(* IEC 61131-3 sources: daoli-st-library/DL_Process (part 14) *)

(* ---- FC_DL_LyoCollapseTempMarginCalc.st ---- *)
(*
  Name: FC_DL_LyoCollapseTempMarginCalc
  Category: DL_Process
  Version: 1.0.0
  Round: R91 / 2026-11-25
  开源溯源：clean-room 自研（族 制药冻干真空冷冻干燥，ST 开源生态实测 0 命中，无外部代码引入）
  功能：1) 塌陷温度裕度 = 塌陷温度 − 制品温度，即 fMarginK = fCollapseC − fProductC，
           裕度为正表示制品温度仍低于塌陷温度（安全侧），为负表示已越过塌陷边界。
        2) 裕度分级（nGrade）：0 = 合格（裕度 >= fMarginWarnK），1 = 预警（fMarginMinK <= 裕度 < fMarginWarnK），
           2 = 不足（裕度 < fMarginMinK），分级判据全部对原始裕度做，钳制只作用于输出数值。
        3) 冰点约束：制品温度必须低于冰点 fIcePointC，否则一次干燥已进入液态（融冰），
           输出 xAboveIce 供上层立即降温或转二次干燥。
  边界条件：1) 非有限值闸：五路实值入参先过 NOT(x > -DL_BIG AND x < DL_BIG)，同时拦 NaN 与 Inf，
           命中即闸断实值通路（裕度强制 0.0 且置分级 2 = 不足），不得只置标志（R19）。
        2) 阈值域闸：分级阈值须满足 fMarginMinK < fMarginWarnK（否则两级判据区间为空、分级恒失效），
           越域判无效并把 nGrade 置 2（保守侧）。
        3) 温度域闸：三路温度必须落在 [-DL_T_SPAN, +DL_T_SPAN] 内，越域判无效（量级异常）。
        4) 判据取原始值（R24）：分级与冰点判定使用原始入参，不先把温度夹到工艺带再判。
        5) 物理域钳制：裕度钳到 [-DL_MARGIN_SPAN, +DL_MARGIN_SPAN]，避免极端值污染显示与趋势。
        6) 纯函数无状态：分级不做迟滞，防抖与联锁延时由搁板温控 FB 承担。
  量纲自证：fMarginK = (degC) − (degC) = (K)；与 fMarginMinK / fMarginWarnK 同为温差点量纲 [K]，
           可与温差阈值直接比较；nGrade 为无量纲等级 [level]。
  修订历史 Revision :
    2026-11-25  v1.0.0  R91 首版
*)

FUNCTION FC_DL_LyoCollapseTempMarginCalc : BOOL
VAR_INPUT
    fProductC        : REAL;   // 制品（瓶内）温度 [degC] / Product temperature inside the vial [degC]
    fCollapseC       : REAL;   // 配方给出的塌陷温度 [degC] / Formulation collapse temperature [degC]
    fIcePointC       : REAL;   // 配方给出的冰点 [degC] / Formulation ice point [degC]
    fMarginMinK      : REAL;   // 裕度不足阈值（低于即判不足）[K] / Margin insufficient threshold [K]
    fMarginWarnK     : REAL;   // 裕度预警阈值（低于即判预警）[K] / Margin warning threshold [K]
END_VAR
VAR_OUTPUT
    fMarginK         : REAL;   // 塌陷温度裕度 [K] / Collapse temperature margin [K]
    nGrade           : INT;    // 裕度分级 0=合格 1=预警 2=不足 [level] / Margin grade 0/1/2 [level]
    xMarginLow       : BOOL;   // 裕度不足标志（< 下限）[bool] / Margin insufficient flag [bool]
    xAboveIce        : BOOL;   // 制品温度高于冰点标志 [bool] / Product above ice point flag [bool]
    xValid           : BOOL;   // 计算有效标志 [bool] / Calculation valid flag [bool]
END_VAR
VAR
    _fMarginRawK     : REAL;   // 钳制前的原始裕度 [K] / Raw margin before limiting [K]
END_VAR
VAR CONSTANT
    DL_BIG           : REAL := 1.0E12;    // 非有限值闸量级上限 [-] / Finiteness gate magnitude [-]
    DL_EPS           : REAL := 1.0E-9;    // 数值零闸阈值 [-] / Numeric zero gate threshold [-]
    DL_T_SPAN        : REAL := 300.0;     // 温度量级闸跨度 [degC] / Temperature magnitude gate span [degC]
    DL_MARGIN_SPAN   : REAL := 200.0;     // 裕度钳制跨度 [K] / Margin clamp span [K]
    DL_GRADE_OK      : INT := 0;          // 分级：合格 [level] / Grade: acceptable [level]
    DL_GRADE_WARN    : INT := 1;          // 分级：预警 [level] / Grade: warning [level]
    DL_GRADE_BAD     : INT := 2;          // 分级：不足 [level] / Grade: insufficient [level]
END_VAR

(* —— 段 1：非有限值闸（R19：闸断实值通路；失效侧分级置不足） —— *)
IF NOT (fProductC > -DL_BIG AND fProductC < DL_BIG)
   OR NOT (fCollapseC > -DL_BIG AND fCollapseC < DL_BIG)
   OR NOT (fIcePointC > -DL_BIG AND fIcePointC < DL_BIG)
   OR NOT (fMarginMinK > -DL_BIG AND fMarginMinK < DL_BIG)
   OR NOT (fMarginWarnK > -DL_BIG AND fMarginWarnK < DL_BIG) THEN
    fMarginK := 0.0;                        // 输出强制 0.0，切断污染源 / Force zero, cut polluted path
    nGrade := DL_GRADE_BAD;                 // 失效侧按不足处理（保守侧）/ Treat as insufficient when invalid
    xMarginLow := TRUE;                     // 失效侧不足位置真（保守侧）/ Insufficient flag true when invalid
    xAboveIce := FALSE;                     // 失效侧冰点位保持假 / Ice-point flag stays false
    xValid := FALSE;                        // 有效位清零 / Validity cleared
    FC_DL_LyoCollapseTempMarginCalc := FALSE;   // 返回码与有效位同源 / Return mirrors validity
    RETURN;                                 // 立即退出 / Immediate exit
END_IF

(* —— 段 2：主算式（不钳制，先出原始值供段 3 判据使用，R24） —— *)
_fMarginRawK := fCollapseC - fProductC;                                           // 塌陷温度裕度 [K]

(* —— 段 3：判据与分级（全部取原始值；单点 BOOL 聚合避免多处赋 FALSE 覆盖） —— *)
xMarginLow := (_fMarginRawK < fMarginMinK);                                       // 裕度不足
xAboveIce := (fProductC > fIcePointC);                                            // 已融冰（高于冰点）
xValid := (fMarginMinK < fMarginWarnK)                                            // 分级阈值必须有效（min < warn）
          AND (ABS(fProductC) <= DL_T_SPAN)                                       // 温度量级闸
          AND (ABS(fCollapseC) <= DL_T_SPAN)
          AND (ABS(fIcePointC) <= DL_T_SPAN)
          AND (fCollapseC > fIcePointC);                                          // 塌陷温度须高于冰点（物理约束）

IF NOT xValid THEN
    nGrade := DL_GRADE_BAD;                 // 参数非法：按不足处理（保守侧）
ELSIF _fMarginRawK >= fMarginWarnK THEN
    nGrade := DL_GRADE_OK;                  // 裕度充足
ELSIF _fMarginRawK >= fMarginMinK THEN
    nGrade := DL_GRADE_WARN;                // 预警带
ELSE
    nGrade := DL_GRADE_BAD;                 // 不足
END_IF

(* —— 段 4：输出单点写盘（钳制到物理域内，分级已在段 3 定案） —— *)
fMarginK := LIMIT(-DL_MARGIN_SPAN, _fMarginRawK, DL_MARGIN_SPAN);                  // 裕度钳到物理域 [K]
FC_DL_LyoCollapseTempMarginCalc := xValid;                                        // 返回码：TRUE = 计算可信

END_FUNCTION

(* ---- FC_DL_LyoIceVaporPressureCalc.st ---- *)
(*
  Name: FC_DL_LyoIceVaporPressureCalc
  Category: DL_Process
  Version: 1.0.0
  Round: R91 / 2026-11-25
  开源溯源：clean-room 自研（族 制药冻干真空冷冻干燥，ST 开源生态实测 0 命中，无外部代码引入）
  功能：1) 冰面饱和蒸气压按 Magnus 型 Goff-Gratch 简化式求解：
           p_ice = 611.15 * EXP(22.452 * T / (272.55 + T))，T 为冰面温度 [degC]，
           611.15 为 0 degC 时冰面饱和蒸气压 [Pa]，22.452 与 272.55 为冰相经验常数。
           该式在 -60 ~ 0 degC 内相对误差小于 1 %，是冻干一次干燥压力设定的标准依据。
        2) 派生输出过冷度裕量 fSubcoolK = 0.0 − T，即离冰点的距离；
           冻干工艺要求制品温度始终低于冰点，裕量为负意味着已融冰（塌陷前兆）。
        3) 温度域校验：温度必须落在 [DL_T_LO, DL_T_HI] = [-60.0, 0.0] degC 内，
           越域只置 xDomainOk = FALSE 而数值钳到域内输出，因为经验常数在域外已失效。
  边界条件：1) 非有限值闸：温度入参先过 NOT(x > -DL_BIG AND x < DL_BIG)，同时拦 NaN 与 Inf，
           命中即闸断实值通路（fPressurePa 与 fSubcoolK 强制 0.0），不得只置标志（R19）。
        2) 分母零闸：经验式分母 272.55 + T 在 T = -272.55 degC 处为零，
           本件温度域下限 -60 degC 远高于该点，但仍显式校验 |272.55 + T| > DL_EPS，
           防止越域调用（下游误传开尔文值）导致除零。
        3) 指数溢出闸：指数 22.452*T/(272.55+T) 在接近 -272.55 时发散，
           计算前用温度域闸先拦截，绝不让 EXP 收到发散指数（EXP 溢出为 Inf 会穿透下游）。
        4) 判据取原始值（R24）：温度越域判定使用原始入参 fTempC，不对其先钳制再判。
        5) 物理域钳制：气压钳 0.0 ~ DL_P_HI_PA；过冷度钳到 [-DL_T_HI_SPAN, +DL_T_HI_SPAN]。
        6) 纯函数无状态：不做滤波，测点噪声抑制由下游一阶滤波件承担。
  量纲自证：T [degC] 代入经验式时以温差形式参与（degC 与 K 的差值尺度相同），
           22.452*T/(272.55+T) = (无因次)，故 EXP 的自变量无因次；
           p_ice = (Pa) * (无因次) = Pa，量纲合法。
  修订历史 Revision :
    2026-11-25  v1.0.0  R91 首版
*)

FUNCTION FC_DL_LyoIceVaporPressureCalc : BOOL
VAR_INPUT
    fTempC           : REAL;   // 冰面温度 [degC] / Ice surface temperature [degC]
END_VAR
VAR_OUTPUT
    fPressurePa      : REAL;   // 冰面饱和蒸气压 [Pa] / Ice surface saturation vapour pressure [Pa]
    fSubcoolK        : REAL;   // 距冰点的过冷度裕量 [K] / Subcooling margin below the ice point [K]
    xDomainOk        : BOOL;   // 温度在经验式有效域内 [bool] / Temperature within the valid domain [bool]
    xValid           : BOOL;   // 计算有效标志 [bool] / Calculation valid flag [bool]
END_VAR
VAR
    _fDenomK         : REAL;   // 经验式分母（272.55 + T）[K] / Empirical denominator, 272.55 + T [K]
    _fExpo           : REAL;   // 经验式指数（无因次）[-] / Empirical exponent, dimensionless [-]
    _fPressRawPa     : REAL;   // 钳制前的原始气压 [Pa] / Raw pressure before limiting [Pa]
    _fTempUseC       : REAL;   // 域钳制后参与计算的温度 [degC] / Temperature used after domain clamping [degC]
END_VAR
VAR CONSTANT
    DL_EPS           : REAL := 1.0E-9;    // 数值零闸阈值 [-] / Numeric zero gate threshold [-]
    DL_BIG           : REAL := 1.0E12;    // 非有限值闸量级上限 [-] / Finiteness gate magnitude [-]
    DL_T_LO          : REAL := -60.0;     // 经验式有效温度下限 [degC] / Valid temperature low bound [degC]
    DL_T_HI          : REAL := 0.0;       // 经验式有效温度上限（冰点）[degC] / Valid temperature high, ice point [degC]
    DL_P0_PA         : REAL := 611.15;    // 0 degC 冰面饱和蒸气压 [Pa] / Ice saturation pressure at 0 degC [Pa]
    DL_COEF_A        : REAL := 22.452;    // 冰相经验常数 A（无因次）[-] / Ice-phase empirical constant A [-]
    DL_COEF_B        : REAL := 272.55;    // 冰相经验常数 B [K] / Ice-phase empirical constant B [K]
    DL_P_HI_PA       : REAL := 700.0;     // 气压物理上限（略高于 0 degC 冰面值）[Pa] / Pressure upper bound [Pa]
    DL_MARGIN_SPAN   : REAL := 200.0;     // 过冷度裕量钳制跨度 [K] / Subcooling margin clamp span [K]
END_VAR

(* —— 段 1：非有限值闸（R19：闸断实值通路） —— *)
IF NOT (fTempC > -DL_BIG AND fTempC < DL_BIG) THEN
    fPressurePa := 0.0;                     // 输出强制 0.0，切断污染源 / Force zero, cut polluted path
    fSubcoolK := 0.0;                       // 裕量强制 0.0 / Margin forced to zero
    xDomainOk := FALSE;                     // 域位清零 / Domain flag cleared
    xValid := FALSE;                        // 有效位清零 / Validity cleared
    FC_DL_LyoIceVaporPressureCalc := FALSE; // 返回码与有效位同源 / Return mirrors validity
    RETURN;                                 // 立即退出 / Immediate exit
END_IF

(* —— 段 2：判据取原始值（R24：先判域，再钳制，禁先钳后判） —— *)
xDomainOk := (fTempC >= DL_T_LO) AND (fTempC <= DL_T_HI);

(* —— 段 3：域钳制后参与计算（经验常数在域外失效，绝不让 EXP 收到发散指数） —— *)
_fTempUseC := LIMIT(DL_T_LO, fTempC, DL_T_HI);                          // 温度钳到有效域 [degC]
_fDenomK := DL_COEF_B + _fTempUseC;                                     // 经验式分母 [K]

(* —— 段 4：分母零闸（防越域调用传开尔文值导致除零，R4） —— *)
IF ABS(_fDenomK) <= DL_EPS THEN
    fPressurePa := 0.0;                     // 分母为零即不可算 / No denominator, no result
    fSubcoolK := 0.0;                       // 裕量不可算 / Margin not computable
    xDomainOk := FALSE;                     // 判域外 / Out of domain
    xValid := FALSE;                        // 判无效 / Invalid
    FC_DL_LyoIceVaporPressureCalc := FALSE; // 返回码同步 / Return synchronised
    RETURN;                                 // 提前退出 / Early exit
END_IF

(* —— 段 5：主算式（Goff-Gratch 简化式，指数自变量已由段 3 钳制保证有界） —— *)
_fExpo := DL_COEF_A * _fTempUseC / _fDenomK;                            // 指数（无因次）[-]
_fPressRawPa := DL_P0_PA * EXP(_fExpo);                                 // 冰面饱和蒸气压 [Pa]
fSubcoolK := LIMIT(-DL_MARGIN_SPAN, DL_T_HI - _fTempUseC, DL_MARGIN_SPAN);   // 过冷度裕量 [K]

(* —— 段 6：输出单点写盘（气压钳制到物理域；有限性已由段 1 保证） —— *)
fPressurePa := LIMIT(0.0, _fPressRawPa, DL_P_HI_PA);                    // 气压钳 0..物理上限 [Pa]
xValid := xDomainOk AND (fPressurePa > 0.0);                            // 域内且有正压才算有效
FC_DL_LyoIceVaporPressureCalc := xValid;                                // 返回码：TRUE = 计算可信

END_FUNCTION

(* ---- FC_DL_LyoPrimaryDryingTimeCalc.st ---- *)
(*
  Name: FC_DL_LyoPrimaryDryingTimeCalc
  Category: DL_Process
  Version: 1.0.0
  Round: R91 / 2026-11-25
  开源溯源：clean-room 自研（族 制药冻干真空冷冻干燥，ST 开源生态实测 0 命中，无外部代码引入）
  功能：1) 一次干燥时间按「可去除水量 / 升华速率」估算：
           可去除水量 W = 装量质量 * (初始含水率 − 目标含水率) / 100，单位 kg；
           时间 t = W / rate，单位 h；rate 为该批量的实测升华速率 [kg/h]。
        2) 水量守恒校验：目标含水率必须低于初始含水率，否则水量为负（配方错），
           判无效而不取绝对值 —— 负水量意味着「越干越湿」的错误配方。
        3) 收敛判据：估算时间超过 fMaxTimeH（工艺允许最长一次干燥时间）时置 xNotConverge，
           表示按当前速率无法在允许时间内达到目标含水率，需提高搁板温度或降低装量。
  边界条件：1) 非有限值闸：五路实值入参先过 NOT(x > -DL_BIG AND x < DL_BIG)，同时拦 NaN 与 Inf，
           命中即闸断实值通路（时间与水量强制 0.0），不得只置标志（R19）。
        2) 速率零闸：升华速率 fRateKgh 必须 > DL_EPS（时间式的分母），否则判无效并清零，
           不得输出「无穷长时间」这种不可执行值。
        3) 含水率域闸：初始与目标含水率必须落在 [0.0, 100.0] % 内，
           装量质量须 > DL_EPS；任一越域判无效，不做钳制。
        4) 判据取原始值（R24）：不收敛判定使用钳制前的 _fTimeRawH，不得先钳再判。
        5) 物理域钳制：时间钳 0.0 ~ DL_TIME_HI_H；水量钳 0.0 ~ 装量质量（水量不可能大于装量）。
        6) 纯函数无状态：不累计已干燥时间，累计与阶段切换由干燥序 FB 承担。
  量纲自证：W = (kg) * (无因次百分数/100) = kg；
           t = (kg)/(kg/h) = h，与 fMaxTimeH 同量纲 [h]，可直接比较。
  修订历史 Revision :
    2026-11-25  v1.0.0  R91 首版
*)

FUNCTION FC_DL_LyoPrimaryDryingTimeCalc : BOOL
VAR_INPUT
    fFillMassKg      : REAL;   // 单批装量质量 [kg] / Batch fill mass [kg]
    fInitMoistPct    : REAL;   // 初始含水率 [%] / Initial moisture content [%]
    fTargetMoistPct  : REAL;   // 目标含水率 [%] / Target moisture content [%]
    fRateKgh         : REAL;   // 该批量实测升华速率 [kg/h] / Measured batch sublimation rate [kg/h]
    fMaxTimeH        : REAL;   // 工艺允许最长一次干燥时间 [h] / Permitted maximum primary drying time [h]
END_VAR
VAR_OUTPUT
    fTimeH           : REAL;   // 一次干燥估算时间 [h] / Estimated primary drying time [h]
    fWaterKg         : REAL;   // 需去除水量 [kg] / Water mass to be removed [kg]
    xNotConverge     : BOOL;   // 超允许时间标志（不收敛）[bool] / Non-convergence flag [bool]
    xValid           : BOOL;   // 计算有效标志 [bool] / Calculation valid flag [bool]
END_VAR
VAR
    _fWaterRawKg     : REAL;   // 钳制前的原始水量 [kg] / Raw water mass before limiting [kg]
    _fTimeRawH       : REAL;   // 钳制前的原始时间 [h] / Raw time before limiting [h]
END_VAR
VAR CONSTANT
    DL_EPS           : REAL := 1.0E-9;    // 数值零闸阈值 [-] / Numeric zero gate threshold [-]
    DL_BIG           : REAL := 1.0E12;    // 非有限值闸量级上限 [-] / Finiteness gate magnitude [-]
    DL_PCT           : REAL := 100.0;     // 百分比换算因子（含水率分母）[%] / Percent conversion factor [%]
    DL_PCT_HI        : REAL := 100.0;     // 含水率物理上限 [%] / Moisture content upper bound [%]
    DL_TIME_HI_H     : REAL := 10000.0;   // 时间物理上限 [h] / Time physical upper bound [h]
END_VAR

(* —— 段 1：非有限值闸（R19：闸断实值通路） —— *)
IF NOT (fFillMassKg > -DL_BIG AND fFillMassKg < DL_BIG)
   OR NOT (fInitMoistPct > -DL_BIG AND fInitMoistPct < DL_BIG)
   OR NOT (fTargetMoistPct > -DL_BIG AND fTargetMoistPct < DL_BIG)
   OR NOT (fRateKgh > -DL_BIG AND fRateKgh < DL_BIG)
   OR NOT (fMaxTimeH > -DL_BIG AND fMaxTimeH < DL_BIG) THEN
    fTimeH := 0.0;                          // 输出强制 0.0，切断污染源 / Force zero, cut polluted path
    fWaterKg := 0.0;                        // 水量强制 0.0 / Water mass forced to zero
    xNotConverge := TRUE;                   // 失效侧按不收敛处理（安全侧）/ Treat as non-converged when invalid
    xValid := FALSE;                        // 有效位清零 / Validity cleared
    FC_DL_LyoPrimaryDryingTimeCalc := FALSE;   // 返回码与有效位同源 / Return mirrors validity
    RETURN;                                 // 立即退出 / Immediate exit
END_IF

(* —— 段 2：分母零闸与域闸（时间式分母为速率；含水率须在 0~100 %） —— *)
IF (fRateKgh <= DL_EPS)                                           // 速率不可为零
   OR (fFillMassKg <= DL_EPS)                                     // 装量不可为零
   OR (fInitMoistPct < 0.0)                                       // 含水率不得为负
   OR (fInitMoistPct > DL_PCT_HI)                                 // 含水率不得超 100 %
   OR (fTargetMoistPct < 0.0)                                     // 目标含水率不得为负
   OR (fTargetMoistPct > DL_PCT_HI)                               // 目标含水率不得超 100 %
   OR (fMaxTimeH <= DL_EPS) THEN                                  // 允许时间必须已组态
    fTimeH := 0.0;                          // 参数不可用即无时间 / No parameter, no time
    fWaterKg := 0.0;                        // 水量不可算 / Water mass not computable
    xNotConverge := TRUE;                   // 按不收敛处理 / Treat as non-converged
    xValid := FALSE;                        // 判无效 / Invalid
    FC_DL_LyoPrimaryDryingTimeCalc := FALSE;   // 返回码同步 / Return synchronised
    RETURN;                                 // 提前退出 / Early exit
END_IF

(* —— 段 3：主算式（不钳制，先出原始值供段 4 判据使用，R24） —— *)
_fWaterRawKg := fFillMassKg * (fInitMoistPct - fTargetMoistPct) / DL_PCT;          // 需去除水量 [kg]
_fTimeRawH := _fWaterRawKg / fRateKgh;                                            // 估算时间 [h]

(* —— 段 4：判据（取原始值；单点 BOOL 聚合避免多处赋 FALSE 覆盖） —— *)
xNotConverge := (_fTimeRawH > fMaxTimeH);                                         // 超允许时间：不收敛
xValid := (_fWaterRawKg >= 0.0)                                                   // 水量不得为负（配方方向固定）
          AND (_fTimeRawH >= 0.0)                                                 // 时间不得为负
          AND (fMaxTimeH <= DL_TIME_HI_H)                                         // 允许时间不得超物理上限
          AND (fInitMoistPct > fTargetMoistPct);                                  // 初始必须高于目标（方向固定）

(* —— 段 5：输出单点写盘（钳制到物理域内，判定结果已在段 4 定案） —— *)
fWaterKg := LIMIT(0.0, _fWaterRawKg, fFillMassKg);                                // 水量钳 0..装量 [kg]
fTimeH := LIMIT(0.0, _fTimeRawH, DL_TIME_HI_H);                                   // 时间钳 0..物理上限 [h]
FC_DL_LyoPrimaryDryingTimeCalc := xValid;                                         // 返回码：TRUE = 计算可信

END_FUNCTION

(* ---- FC_DL_LyoResidualMoistureCalc.st ---- *)
(*
  Name: FC_DL_LyoResidualMoistureCalc
  Category: DL_Process
  Version: 1.0.0
  Round: R91 / 2026-11-25
  开源溯源：clean-room 自研（族 制药冻干真空冷冻干燥，ST 开源生态实测 0 命中，无外部代码引入）
  功能：1) 残余水分估算按「压力升速率法」：一次干燥末期关闭隔离阀，测腔内压力升幅与时间，
           升压速率 r = dP / t [mbar/s]；残余水分与升压速率近似成正比，并用干重比归一：
           W_res% = coef * r / ratio，coef 为经方法学验证的标定系数 [%*s/mbar]，
           ratio 为干物质质量占比 [kg/kg]（干重比），用于把腔体自由水折算到制品含湿量。
        2) 合格判据：残余水分 <= fSpecMaxPct（药典/内控限度，通常 1~3 %）输出 xSpecOver = FALSE。
        3) 比值域校验：干重比必须落在 (DL_RATIO_LO, 1.0] 内（干物质不可能超过总质量，
           也不可能为零），越域判无效而非钳制 —— 钳制会严重放大或抹平结果。
  边界条件：1) 非有限值闸：五路实值入参先过 NOT(x > -DL_BIG AND x < DL_BIG)，同时拦 NaN 与 Inf，
           命中即闸断实值通路（水分与速率强制 0.0 且置超限位，保守侧），不得只置标志（R19）。
        2) 时间零闸：升压时长 fRiseTimeS 必须 > DL_EPS（速率式分母），否则判无效。
        3) 比值零闸：干重比 fDryWeightRatio 必须 > DL_RATIO_LO（水分式分母），否则判无效。
        4) 标定系数域闸：fCoefPctSPerMbar 必须 > DL_EPS（系数未标定则结果无意义）。
        5) 判据取原始值（R24）：超限判定使用钳制前的 _fResRawPct，不得先钳再判。
        6) 物理域钳制：残余水分钳 0.0 ~ DL_PCT_HI；升压速率钳 0.0 ~ DL_RATE_HI。
  量纲自证：r = (mbar)/(s) = mbar/s；
           coef * r / ratio = (%*s/mbar)*(mbar/s)/(kg/kg) = %，干重比无因次，量纲链闭合。
  修订历史 Revision :
    2026-11-25  v1.0.0  R91 首版
*)

FUNCTION FC_DL_LyoResidualMoistureCalc : BOOL
VAR_INPUT
    fPressRiseMbar   : REAL;   // 测试期腔内压力升幅 [mbar] / Chamber pressure rise during the test [mbar]
    fRiseTimeS       : REAL;   // 升压时长 [s] / Pressure rise duration [s]
    fDryWeightRatio  : REAL;   // 干物质质量占比（干重比）[kg/kg] / Dry matter mass ratio [kg/kg]
    fCoefPctSPerMbar : REAL;   // 标定系数 [%*s/mbar] / Calibration coefficient [%*s/mbar]
    fSpecMaxPct      : REAL;   // 残余水分内控上限 [%] / In-house residual moisture limit [%]
END_VAR
VAR_OUTPUT
    fResidualPct     : REAL;   // 估算残余水分 [%] / Estimated residual moisture [%]
    fRiseRateMbarS   : REAL;   // 压力升速率 [mbar/s] / Pressure rise rate [mbar/s]
    xSpecOver        : BOOL;   // 超内控上限标志 [bool] / Over-specification flag [bool]
    xValid           : BOOL;   // 计算有效标志 [bool] / Calculation valid flag [bool]
END_VAR
VAR
    _fRateRawMbarS   : REAL;   // 钳制前的原始升压速率 [mbar/s] / Raw rise rate before limiting [mbar/s]
    _fResRawPct      : REAL;   // 钳制前的原始残余水分 [%] / Raw residual moisture before limiting [%]
END_VAR
VAR CONSTANT
    DL_EPS           : REAL := 1.0E-9;    // 数值零闸阈值 [-] / Numeric zero gate threshold [-]
    DL_BIG           : REAL := 1.0E12;    // 非有限值闸量级上限 [-] / Finiteness gate magnitude [-]
    DL_PCT           : REAL := 100.0;     // 百分比换算因子 [%] / Percent conversion factor [%]
    DL_RATIO_LO      : REAL := 1.0E-6;    // 干重比下限阈值 [kg/kg] / Dry-weight ratio low gate [kg/kg]
    DL_RATIO_HI      : REAL := 1.0;       // 干重比物理上限 [kg/kg] / Dry-weight ratio upper bound [kg/kg]
    DL_RATE_HI       : REAL := 100.0;     // 升压速率物理上限 [mbar/s] / Rise rate upper bound [mbar/s]
END_VAR

(* —— 段 1：非有限值闸（R19：闸断实值通路；失效侧超限位置真，保守侧） —— *)
IF NOT (fPressRiseMbar > -DL_BIG AND fPressRiseMbar < DL_BIG)
   OR NOT (fRiseTimeS > -DL_BIG AND fRiseTimeS < DL_BIG)
   OR NOT (fDryWeightRatio > -DL_BIG AND fDryWeightRatio < DL_BIG)
   OR NOT (fCoefPctSPerMbar > -DL_BIG AND fCoefPctSPerMbar < DL_BIG)
   OR NOT (fSpecMaxPct > -DL_BIG AND fSpecMaxPct < DL_BIG) THEN
    fResidualPct := 0.0;                    // 输出强制 0.0，切断污染源 / Force zero, cut polluted path
    fRiseRateMbarS := 0.0;                  // 速率强制 0.0 / Rate forced to zero
    xSpecOver := TRUE;                      // 失效侧按超限处理（保守侧）/ Treat as over-spec when invalid
    xValid := FALSE;                        // 有效位清零 / Validity cleared
    FC_DL_LyoResidualMoistureCalc := FALSE; // 返回码与有效位同源 / Return mirrors validity
    RETURN;                                 // 立即退出 / Immediate exit
END_IF

(* —— 段 2：分母零闸与域闸（时长与干重比均为分母；标定系数须已标定） —— *)
IF (fRiseTimeS <= DL_EPS)                                         // 时长不可为零
   OR (fDryWeightRatio <= DL_RATIO_LO)                            // 干重比不可为零
   OR (fDryWeightRatio > DL_RATIO_HI)                             // 干重比不得超过 1
   OR (fCoefPctSPerMbar <= DL_EPS)                                // 标定系数必须为正
   OR (fSpecMaxPct <= DL_EPS)                                     // 内控上限必须已组态
   OR (fPressRiseMbar < 0.0) THEN                                 // 升幅不得为负（隔离后压力只升）
    fResidualPct := 0.0;                    // 参数不可用即无结果 / No parameter, no result
    fRiseRateMbarS := 0.0;                  // 速率不可算 / Rate not computable
    xSpecOver := TRUE;                      // 按超限处理（保守侧）/ Treat as over-spec
    xValid := FALSE;                        // 判无效 / Invalid
    FC_DL_LyoResidualMoistureCalc := FALSE; // 返回码同步 / Return synchronised
    RETURN;                                 // 提前退出 / Early exit
END_IF

(* —— 段 3：主算式（不钳制，先出原始值供段 4 判据使用，R24） —— *)
_fRateRawMbarS := fPressRiseMbar / fRiseTimeS;                                    // 升压速率 [mbar/s]
_fResRawPct := fCoefPctSPerMbar * _fRateRawMbarS / fDryWeightRatio;               // 残余水分 [%]

(* —— 段 4：判据（取原始值；单点 BOOL 聚合避免多处赋 FALSE 覆盖） —— *)
xSpecOver := (_fResRawPct > fSpecMaxPct);                                         // 超内控上限
xValid := (_fResRawPct >= 0.0)                                                    // 水分不得为负
          AND (_fResRawPct <= DL_PCT)                                             // 水分不得超过 100 %（量级闸）
          AND (_fRateRawMbarS <= DL_RATE_HI);                                     // 速率不得超物理上限

(* —— 段 5：输出单点写盘（钳制到物理域内，判定结果已在段 4 定案） —— *)
fResidualPct := LIMIT(0.0, _fResRawPct, DL_PCT);                                  // 水分钳 0..100 [%]
fRiseRateMbarS := LIMIT(0.0, _fRateRawMbarS, DL_RATE_HI);                          // 速率钳 0..物理上限 [mbar/s]
FC_DL_LyoResidualMoistureCalc := xValid;                                          // 返回码：TRUE = 计算可信

END_FUNCTION

(* ---- FC_DL_LyoShelfHeatDutyCalc.st ---- *)
(*
  Name: FC_DL_LyoShelfHeatDutyCalc
  Category: DL_Process
  Version: 1.0.0
  Round: R91 / 2026-11-25
  开源溯源：clean-room 自研（族 制药冻干真空冷冻干燥，ST 开源生态实测 0 命中，无外部代码引入）
  功能：1) 搁板加热功率按「升华吸热 / 加热效率」计算：
           P = rate * latent / eff / 3600，rate 为升华速率 [kg/h]、latent 为升华潜热 [kJ/kg]，
           3600 为 kJ/h 到 kW 的时基折算；eff 为搁板到制品的综合传热效率。
           该功率是一次干燥期搁板温度控制器的前馈给定。
        2) 功率负荷率 fDutyLoadPct = P / fHeaterMaxKw * 100，用于判断是否已触及加热器额定上限；
           超上限只置 xDutyOver 并钳到额定值，不把越限值当作可执行指令下发。
        3) 效率物理域校验：eff 必须落在 (0.0, 1.0] 内，大于 1 违反热力学第一定律，
           视为组态错误判无效（不钳制，钳制会把非法组态伪装成合法）。
  边界条件：1) 非有限值闸：四路实值入参先过 NOT(x > -DL_BIG AND x < DL_BIG)，同时拦 NaN 与 Inf，
           命中即闸断实值通路（功率与负荷率强制 0.0），不得只置标志（R19）。
        2) 分母零闸：加热效率 fHeatEff 与加热器额定功率 fHeaterMaxKw 均须 > DL_EPS，
           否则功率式与负荷率式分母为零，直接判无效。
        3) 潜热域闸：升华潜热 fLatentKjKg 必须落在 (DL_LATENT_LO, DL_LATENT_HI) 内，
           越域说明工质不是水（冰的升华潜热约 2838 kJ/kg），判无效以免误算他物质。
        4) 判据取原始值（R24）：超上限判定使用钳制前的 _fDutyRawKw，不得先钳再判。
        5) 物理域钳制：功率钳 0.0 ~ fHeaterMaxKw；负荷率钳 0.0 ~ DL_PCT_HI。
        6) 纯函数无状态：不做功率限幅斜坡，斜坡由搁板温控 FB 承担。
  量纲自证：rate [kg/h] * latent [kJ/kg] = (kJ/h)；除以 3600 (s/h) 得 kJ/s = kW；
           再除以无因次效率 eff 仍为 kW，与 fHeaterMaxKw 同量纲；
           fDutyLoadPct = (kW)/(kW)*100 = 无因次百分数 [%]，量纲合法。
  修订历史 Revision :
    2026-11-25  v1.0.0  R91 首版
*)

FUNCTION FC_DL_LyoShelfHeatDutyCalc : BOOL
VAR_INPUT
    fRateKgh         : REAL;   // 升华速率 [kg/h] / Sublimation rate [kg/h]
    fLatentKjKg      : REAL;   // 升华潜热 [kJ/kg] / Latent heat of sublimation [kJ/kg]
    fHeatEff         : REAL;   // 搁板到制品综合传热效率（0~1 无因次）[-] / Shelf-to-product heat efficiency [-]
    fHeaterMaxKw     : REAL;   // 搁板加热器额定功率 [kW] / Rated shelf heater power [kW]
END_VAR
VAR_OUTPUT
    fDutyKw          : REAL;   // 所需加热功率 [kW] / Required heating duty [kW]
    fDutyLoadPct     : REAL;   // 加热功率负荷率 [%] / Heating duty load ratio [%]
    xDutyOver        : BOOL;   // 功率超额定标志 [bool] / Duty overrun flag [bool]
    xValid           : BOOL;   // 计算有效标志 [bool] / Calculation valid flag [bool]
END_VAR
VAR
    _fDutyRawKw      : REAL;   // 钳制前的原始功率 [kW] / Raw duty before limiting [kW]
    _fLoadRawPct     : REAL;   // 钳制前的原始负荷率 [%] / Raw load ratio before limiting [%]
END_VAR
VAR CONSTANT
    DL_EPS           : REAL := 1.0E-9;    // 数值零闸阈值 [-] / Numeric zero gate threshold [-]
    DL_BIG           : REAL := 1.0E12;    // 非有限值闸量级上限 [-] / Finiteness gate magnitude [-]
    DL_SEC_PER_H     : REAL := 3600.0;    // 小时到秒的时基折算 [s/h] / Seconds per hour [s/h]
    DL_PCT           : REAL := 100.0;     // 百分比换算因子 [%] / Percent conversion factor [%]
    DL_PCT_HI        : REAL := 100.0;     // 负荷率物理上限 [%] / Load ratio upper bound [%]
    DL_EFF_HI        : REAL := 1.0;       // 传热效率物理上限（热力学第一定律）[-] / Efficiency upper bound [-]
    DL_LATENT_LO     : REAL := 2000.0;    // 冰升华潜热域下限 [kJ/kg] / Ice latent heat domain low [kJ/kg]
    DL_LATENT_HI     : REAL := 4000.0;    // 冰升华潜热域上限 [kJ/kg] / Ice latent heat domain high [kJ/kg]
END_VAR

(* —— 段 1：非有限值闸（R19：闸断实值通路） —— *)
IF NOT (fRateKgh > -DL_BIG AND fRateKgh < DL_BIG)
   OR NOT (fLatentKjKg > -DL_BIG AND fLatentKjKg < DL_BIG)
   OR NOT (fHeatEff > -DL_BIG AND fHeatEff < DL_BIG)
   OR NOT (fHeaterMaxKw > -DL_BIG AND fHeaterMaxKw < DL_BIG) THEN
    fDutyKw := 0.0;                         // 输出强制 0.0，切断污染源 / Force zero, cut polluted path
    fDutyLoadPct := 0.0;                    // 负荷率强制 0.0 / Load ratio forced to zero
    xDutyOver := FALSE;                     // 失效侧超限位保持假 / Overrun stays false
    xValid := FALSE;                        // 有效位清零 / Validity cleared
    FC_DL_LyoShelfHeatDutyCalc := FALSE;    // 返回码与有效位同源 / Return mirrors validity
    RETURN;                                 // 立即退出 / Immediate exit
END_IF

(* —— 段 2：分母零闸与域闸（效率、额定功率为分母；潜热须为水冰） —— *)
IF (fHeatEff <= DL_EPS)                                           // 效率不可为零
   OR (fHeatEff > DL_EFF_HI)                                      // 效率不得大于 1
   OR (fHeaterMaxKw <= DL_EPS)                                    // 额定功率必须已组态
   OR (fLatentKjKg <= DL_LATENT_LO)                               // 潜热不得低于冰升华域下限
   OR (fLatentKjKg >= DL_LATENT_HI)                               // 潜热不得高于冰升华域上限
   OR (fRateKgh < 0.0) THEN                                       // 速率不得为负（方向固定）
    fDutyKw := 0.0;                         // 参数不可用即无功率 / No parameter, no duty
    fDutyLoadPct := 0.0;                    // 负荷率不可算 / Load ratio not computable
    xDutyOver := FALSE;                     // 超限位保持假 / Overrun stays false
    xValid := FALSE;                        // 判无效 / Invalid
    FC_DL_LyoShelfHeatDutyCalc := FALSE;    // 返回码同步 / Return synchronised
    RETURN;                                 // 提前退出 / Early exit
END_IF

(* —— 段 3：主算式（不钳制，先出原始值供段 4 判据使用，R24） —— *)
_fDutyRawKw := fRateKgh * fLatentKjKg / fHeatEff / DL_SEC_PER_H;                   // 所需功率 [kW]
_fLoadRawPct := _fDutyRawKw / fHeaterMaxKw * DL_PCT;                               // 负荷率 [%]

(* —— 段 4：判据（取原始值；单点 BOOL 聚合避免多处赋 FALSE 覆盖） —— *)
xDutyOver := (_fDutyRawKw > fHeaterMaxKw);                                        // 功率越额定上限
xValid := (_fDutyRawKw >= 0.0)                                                    // 功率不得为负
          AND (_fLoadRawPct >= 0.0);                                              // 负荷率不得为负

(* —— 段 5：输出单点写盘（钳制到物理域内，判定结果已在段 4 定案） —— *)
fDutyKw := LIMIT(0.0, _fDutyRawKw, fHeaterMaxKw);                                 // 功率钳 0..额定 [kW]
fDutyLoadPct := LIMIT(0.0, _fLoadRawPct, DL_PCT_HI);                              // 负荷率钳 0..100 [%]
FC_DL_LyoShelfHeatDutyCalc := xValid;                                             // 返回码：TRUE = 计算可信

END_FUNCTION

(* ---- FC_DL_LyoSublimationRateCalc.st ---- *)
(*
  Name: FC_DL_LyoSublimationRateCalc
  Category: DL_Process
  Version: 1.0.0
  Round: R91 / 2026-11-25
  开源溯源：clean-room 自研（族 制药冻干真空冷冻干燥，ST 开源生态实测 0 命中，无外部代码引入）
  功能：1) 升华速率按「传质推动力式」计算：dm/dt = K * A * (p_ice − p_chamber)，
           K 为综合传质系数（含边界层与干燥层阻力），A 为升华面积，
           p_ice 为冰面饱和蒸气压、p_chamber 为腔体实测压力；输出单位 kg/h。
        2) 压差负值为失效判据：腔体压力高于冰面饱和压力时不存在升华推动力
           （此时是凝华而非升华），输出 xNoDrive = TRUE 且速率强制 0.0，
           绝不把负速率下发给热负荷件（会把加热变成制冷指令）。
        3) 速率上限保护：速率超过 fRateMaxKgh 只置 xRateOver 并把数值钳到上限，
           用于识别「冰面暴沸/产品飞溅」风险工况。
  边界条件：1) 非有限值闸：五路实值入参先过 NOT(x > -DL_BIG AND x < DL_BIG)，同时拦 NaN 与 Inf，
           命中即闸断实值通路（速率与压差强制 0.0），不得只置标志（R19）。
        2) 系数零闸：传质系数 fMassCoefKghPa 与升华面积 fAreaM2 均须 > DL_EPS，
           任一为零则速率恒为零、时间估算发散，直接判无效而非输出 0。
        3) 压差方向闸：dP = p_ice − p_chamber 必须 > DL_EPS 才允许计算速率；
           零压差（平衡态）与负压差（凝华）一律判 xNoDrive 并清零速率。
        4) 压力域闸：两路压力不得为负（负绝压属传感器错），
           fRateMaxKgh 须 > DL_EPS（上限为零会使钳制把一切速率抹平）。
        5) 判据取原始值（R24）：超上限判定使用钳制前的 _fRateRawKgh，不得先钳再判。
        6) 物理域钳制：速率钳 0.0 ~ fRateMaxKgh；压差钳 0.0 ~ DL_DP_HI_PA。
  量纲自证：K [kg/(m2*h*Pa)] * A [m2] * dP [Pa] = (kg/h)，量纲链闭合；
           fDpPa = (Pa) − (Pa) = Pa，与 K 的分母同量纲。
  修订历史 Revision :
    2026-11-25  v1.0.0  R91 首版
*)

FUNCTION FC_DL_LyoSublimationRateCalc : BOOL
VAR_INPUT
    fIcePressPa      : REAL;   // 冰面饱和蒸气压 [Pa] / Ice surface saturation vapour pressure [Pa]
    fChamberPressPa  : REAL;   // 腔体实测压力 [Pa] / Measured chamber pressure [Pa]
    fMassCoefKghPa   : REAL;   // 综合传质系数 [kg/(m2*h*Pa)] / Overall mass transfer coefficient [kg/(m2*h*Pa)]
    fAreaM2          : REAL;   // 有效升华面积 [m2] / Effective sublimation area [m2]
    fRateMaxKgh      : REAL;   // 允许升华速率上限 [kg/h] / Permitted sublimation rate upper limit [kg/h]
END_VAR
VAR_OUTPUT
    fRateKgh         : REAL;   // 升华速率 [kg/h] / Sublimation rate [kg/h]
    fDpPa            : REAL;   // 传质压差（冰面 − 腔体）[Pa] / Driving pressure difference [Pa]
    xNoDrive         : BOOL;   // 无升华推动力标志（压差 <= 0）[bool] / No driving force flag [bool]
    xRateOver        : BOOL;   // 速率超上限标志 [bool] / Rate overrun flag [bool]
    xValid           : BOOL;   // 计算有效标志 [bool] / Calculation valid flag [bool]
END_VAR
VAR
    _fDpRawPa        : REAL;   // 未钳制的压差 [Pa] / Unclamped pressure difference [Pa]
    _fRateRawKgh     : REAL;   // 钳制前的原始速率 [kg/h] / Raw rate before limiting [kg/h]
END_VAR
VAR CONSTANT
    DL_EPS           : REAL := 1.0E-9;    // 数值零闸阈值 [-] / Numeric zero gate threshold [-]
    DL_BIG           : REAL := 1.0E12;    // 非有限值闸量级上限 [-] / Finiteness gate magnitude [-]
    DL_DP_HI_PA      : REAL := 700.0;     // 压差物理上限 [Pa] / Pressure difference upper bound [Pa]
    DL_RATE_ABS_MAX  : REAL := 1000.0;    // 速率绝对物理上限 [kg/h] / Absolute rate upper bound [kg/h]
END_VAR

(* —— 段 1：非有限值闸（R19：闸断实值通路） —— *)
IF NOT (fIcePressPa > -DL_BIG AND fIcePressPa < DL_BIG)
   OR NOT (fChamberPressPa > -DL_BIG AND fChamberPressPa < DL_BIG)
   OR NOT (fMassCoefKghPa > -DL_BIG AND fMassCoefKghPa < DL_BIG)
   OR NOT (fAreaM2 > -DL_BIG AND fAreaM2 < DL_BIG)
   OR NOT (fRateMaxKgh > -DL_BIG AND fRateMaxKgh < DL_BIG) THEN
    fRateKgh := 0.0;                        // 输出强制 0.0，切断污染源 / Force zero, cut polluted path
    fDpPa := 0.0;                           // 压差强制 0.0 / Pressure difference forced to zero
    xNoDrive := TRUE;                       // 失效侧按无推动力处理（安全侧）/ Treat as no drive on invalid
    xRateOver := FALSE;                     // 失效侧超限位保持假 / Overrun stays false
    xValid := FALSE;                        // 有效位清零 / Validity cleared
    FC_DL_LyoSublimationRateCalc := FALSE;  // 返回码与有效位同源 / Return mirrors validity
    RETURN;                                 // 立即退出 / Immediate exit
END_IF

(* —— 段 2：系数零闸（传质系数与面积为乘子，为零则速率恒零、时间估算发散） —— *)
IF (fMassCoefKghPa <= DL_EPS)                                     // 传质系数不可为零
   OR (fAreaM2 <= DL_EPS)                                         // 升华面积不可为零
   OR (fRateMaxKgh <= DL_EPS) THEN                                // 速率上限必须已组态
    fRateKgh := 0.0;                        // 参数不可用即无速率 / No parameter, no rate
    fDpPa := 0.0;                           // 压差不可用 / Difference not usable
    xNoDrive := TRUE;                       // 按无推动力处理 / Treat as no drive
    xRateOver := FALSE;                     // 超限位保持假 / Overrun stays false
    xValid := FALSE;                        // 判无效 / Invalid
    FC_DL_LyoSublimationRateCalc := FALSE;  // 返回码同步 / Return synchronised
    RETURN;                                 // 提前退出 / Early exit
END_IF

(* —— 段 3：压差方向闸（判断据取原始压差，R24） —— *)
_fDpRawPa := fIcePressPa - fChamberPressPa;                        // 传质压差 [Pa]
xNoDrive := (_fDpRawPa <= DL_EPS);                                 // 压差为零或为负：无升华推动力

IF xNoDrive THEN
    fRateKgh := 0.0;                        // 无推动力即零速率（不得下发负速率）
    fDpPa := 0.0;                           // 压差出口钳零 / Difference clamped to zero
    xRateOver := FALSE;                     // 超限位保持假 / Overrun stays false
    xValid := (fIcePressPa >= 0.0) AND (fChamberPressPa >= 0.0);     // 压力非负时计算本身仍可信（平衡态）
    FC_DL_LyoSublimationRateCalc := xValid; // 返回码与有效位同源
    RETURN;                                 // 平衡态/凝华态到此为止 / Stop here for equilibrium or deposition
END_IF

(* —— 段 4：主算式（不钳制，先出原始值供段 5 判据使用） —— *)
_fRateRawKgh := fMassCoefKghPa * fAreaM2 * _fDpRawPa;              // 升华速率 [kg/h]

(* —— 段 5：判据（取原始值；单点 BOOL 聚合避免多处赋 FALSE 覆盖） —— *)
xRateOver := (_fRateRawKgh > fRateMaxKgh);                         // 速率越上限（暴沸/飞溅风险）
xValid := (fIcePressPa >= 0.0)                                     // 压力不得为负（负绝压属传感器错）
          AND (fChamberPressPa >= 0.0)
          AND (fAreaM2 > 0.0)                                      // 面积已验为正
          AND (fRateMaxKgh <= DL_RATE_ABS_MAX)                     // 上限不得超绝对物理上限
          AND (_fRateRawKgh >= 0.0);                               // 速率不得为负（方向固定）

(* —— 段 6：输出单点写盘（钳制到物理域内，判定结果已在段 5 定案） —— *)
fRateKgh := LIMIT(0.0, _fRateRawKgh, fRateMaxKgh);                 // 速率钳 0..工艺上限 [kg/h]
fDpPa := LIMIT(0.0, _fDpRawPa, DL_DP_HI_PA);                       // 压差钳 0..物理上限 [Pa]
FC_DL_LyoSublimationRateCalc := xValid;                            // 返回码：TRUE = 计算可信

END_FUNCTION

(* ---- FC_DL_MashStepInfusionCalc.st ---- *)
// FC_DL_MashStepInfusionCalc v1.0.0
// 开源溯源：clean-room 自研（族 DL_Process，ST 生态实测 0 命中，无外部代码引入）
(*
  功能: 糖化升温热量与蒸汽：Q = m·cp·(T末 − T初)/(1 − 热损率/100) [kJ]，蒸汽 = Q/潜热 [kg]；
        未计入罐体蓄热与投料比热差（工程简化）。
  邻件/码位: 与 FC_DL_WortAerationRateCalc、FC_DL_WortBoilEvaporationCalc 同属前段热工链；
             16#0002_9231 = 非有限、质量/比热/潜热非正、末温不高于初温或热损率越界拒收。
*)
FUNCTION FC_DL_MashStepInfusionCalc : REAL
VAR_INPUT
    fMashMass    : REAL := 5000.0;  // 醪液质量 [kg]，域 > 0 / Mash mass [kg]
    fCp          : REAL := 3.9;     // 醪液比热 [kJ/(kg·K)]，域 > 0 / Specific heat [kJ/(kg K)]
    fTempStart   : REAL := 50.0;    // 升温初温 [°C] / Initial temperature [degC]
    fTempEnd     : REAL := 65.0;    // 升温末温 [°C]，域 > 初温 / Target temperature [degC]
    fLossRate    : REAL := 5.0;     // 热损率 [%]，域 [0, 100) / Heat loss ratio [%]
    fSteamLatent : REAL := 2100.0;  // 蒸汽潜热 [kJ/kg]，域 > 0 / Steam latent heat [kJ/kg]
END_VAR
VAR_OUTPUT
    fHeatNeed  : REAL;              // 需热量 [kJ] / Required heat [kJ]
    fSteamNeed : REAL;              // 需蒸汽量 [kg] / Required steam [kg]
    bValid     : BOOL;              // 结果有效回执 [-] / Result validity receipt
    uErrorId   : UDINT;             // 事件码，0 = 无事件 / Event code
END_VAR
// 段 0：全路径出口安全缺省 / Safe defaults on all outlets
fHeatNeed := 0.0;                   // 需热量缺省零 / Required heat default zero
fSteamNeed := 0.0;                  // 需蒸汽缺省零 / Required steam default zero
bValid := FALSE;                    // 有效回执预清 / Validity preset clear
uErrorId := 16#0000;                // 事件码预清 / Event code preset clear
FC_DL_MashStepInfusionCalc := 0.0;  // 返回值缺省零（镜像需蒸汽）/ Return default zero
// 段 1：非有限闸（六入参全枚举）/ Non-finite gate over all inputs
IF (fMashMass <> fMashMass) OR (fCp <> fCp) OR (fTempStart <> fTempStart)
   OR (fTempEnd <> fTempEnd) OR (fLossRate <> fLossRate) OR (fSteamLatent <> fSteamLatent)
   OR (ABS(fMashMass) >= 3.0E38) OR (ABS(fCp) >= 3.0E38) OR (ABS(fTempStart) >= 3.0E38)
   OR (ABS(fTempEnd) >= 3.0E38) OR (ABS(fLossRate) >= 3.0E38) OR (ABS(fSteamLatent) >= 3.0E38) THEN
    uErrorId := 16#0002_9231;   // 入参非有限拒收 / Non-finite input reject
    RETURN;
END_IF
// 段 2：域闸（质量/比热/潜热为正 + 末温高于初温 + 热损率上界，R4）/ Domain gate
IF (fMashMass <= 1.0E-6) OR (fCp <= 1.0E-6) OR (fSteamLatent <= 1.0E-6) THEN
    uErrorId := 16#0002_9231;   // 质量、比热或潜热非正 / Non-positive mass, capacity or latent
    RETURN;
END_IF
IF fTempEnd <= fTempStart THEN
    uErrorId := 16#0002_9231;   // 末温不高于初温，无需升温 / Target not above initial
    RETURN;
END_IF
IF (fLossRate < 0.0) OR (fLossRate >= 100.0) THEN
    uErrorId := 16#0002_9231;   // 热损率越界（分母近零）/ Heat loss ratio out of range
    RETURN;
END_IF
// 段 3：主计算（需热量 → 需蒸汽）/ Main computation
fHeatNeed := fMashMass * fCp * (fTempEnd - fTempStart) / (1.0 - fLossRate / 100.0);   // 需热量 [kJ]
fSteamNeed := fHeatNeed / fSteamLatent;                         // 需蒸汽 [kg] / Required steam
// 段 4：出口闸（双输出非有限复核 + 正数复核）/ Outlet gate
IF (fHeatNeed <> fHeatNeed) OR (fSteamNeed <> fSteamNeed)
   OR (ABS(fHeatNeed) >= 3.0E38) OR (ABS(fSteamNeed) >= 3.0E38)
   OR (fHeatNeed <= 0.0) OR (fSteamNeed <= 0.0) THEN
    fHeatNeed := 0.0;           // 复核失败回缺省 / Fallback on recheck failure
    fSteamNeed := 0.0;          // 复核失败回缺省 / Fallback on recheck failure
    uErrorId := 16#0002_9231;   // 出口复核拒收 / Output recheck reject
    RETURN;
END_IF
bValid := TRUE;                 // 有效回执 / Validity receipt
FC_DL_MashStepInfusionCalc := fSteamNeed;       // 返回值镜像需蒸汽 / Return mirrors steam demand
END_FUNCTION

(* ---- FC_DL_MashStrikeWaterTempCalc.st ---- *)
(*
  Component : FC_DL_MashStrikeWaterTempCalc
  Category  : DL_Process
  Type      : FC
  Complexity: C2
  VERSION   : v1.0.0
  功能      : 糖化投料水温核算：按麦芽量/比热/初温与水量做能量平衡，反算达到目标醪温所需的投料水温，并含设备热损修正。
  开源溯源  : 道莅原创 clean-room 自研（无外部代码引用）｜License: MIT
  边界条件  : ① 麦芽量、水量、两侧比热均须 > 1e-9，否则返回哨兵 -1（水量热容为除子）；
              ② 热损按目标醪温的百分比上调所需焓，热损率钳位 0~30 %；
              ③ 反算水温可低于 0 °C（需预冷），不下钳位，仅照实输出供上位判断。
*)
FUNCTION FC_DL_MashStrikeWaterTempCalc : REAL
VAR_INPUT
    fMaltKg      : REAL;   (* 麦芽投料量 [kg] Malt charge *)
    fMaltCpKJkgK : REAL;   (* 麦芽比热容 [kJ/(kg·K)] Malt specific heat *)
    fMaltT0C     : REAL;   (* 麦芽初始温度 [°C] Malt initial temperature *)
    fWaterKg     : REAL;   (* 投料水量 [kg] Strike water mass *)
    fWaterCpKJkgK: REAL;   (* 水比热容 [kJ/(kg·K)] Water specific heat *)
    fTargetMashC : REAL;   (* 目标醪液温度 [°C] Target mash temperature *)
    fLossPct     : REAL;   (* 设备热损率 [%] Equipment heat loss ratio *)
END_VAR
VAR_OUTPUT
    fStrikeWaterC : REAL;  (* 所需投料水温 [°C] Required strike water temperature *)
    fHeatCapMaltKJK: REAL; (* 麦芽热容 [kJ/K] Malt heat capacity *)
    fHeatCapWaterKJK: REAL;(* 水热容 [kJ/K] Water heat capacity *)
    xValid        : BOOL;  (* 计算有效性标志 [-] Calculation valid flag *)
END_VAR
VAR CONSTANT
    DL_EPS      : REAL := 1.0E-9;   (* 除零判定容差 [无量纲] Divide-by-zero tolerance *)
    DL_PCT_BASE : REAL := 100.0;    (* 百分比基准 [%] Percent base *)
    DL_LOSS_MAX : REAL := 30.0;     (* 热损率上限 [%] Heat loss upper clamp *)
    DL_ZERO     : REAL := 0.0;      (* 零常量 [无量纲] Zero constant *)
END_VAR
VAR
    fTargetEffC : REAL;   (* 含热损修正的目标温度 [°C] Loss-corrected target temperature *)
    fLossUnit   : REAL;   (* 热损率折算系数 [-] Heat loss as fraction *)
END_VAR
(* 出口预置：四出口统一预置 *)
fStrikeWaterC := 0.0; fHeatCapMaltKJK := 0.0; fHeatCapWaterKJK := 0.0; xValid := FALSE;
(* 非有限拦截：自反判 NaN，自身差值判 Inf *)
IF (fMaltKg <> fMaltKg) OR ((fMaltKg - fMaltKg) <> 0.0)
   OR (fMaltCpKJkgK <> fMaltCpKJkgK) OR ((fMaltCpKJkgK - fMaltCpKJkgK) <> 0.0)
   OR (fMaltT0C <> fMaltT0C) OR ((fMaltT0C - fMaltT0C) <> 0.0)
   OR (fWaterKg <> fWaterKg) OR ((fWaterKg - fWaterKg) <> 0.0)
   OR (fWaterCpKJkgK <> fWaterCpKJkgK) OR ((fWaterCpKJkgK - fWaterCpKJkgK) <> 0.0)
   OR (fTargetMashC <> fTargetMashC) OR ((fTargetMashC - fTargetMashC) <> 0.0)
   OR (fLossPct <> fLossPct) OR ((fLossPct - fLossPct) <> 0.0) THEN
    FC_DL_MashStrikeWaterTempCalc := -1.0;  (* 哨兵 -1：输入非有限 / Sentinel -1 non-finite *)
    RETURN;
END_IF
(* 组态域闸：两侧质量与比热均为比例基，水量热容为除子 *)
IF (fMaltKg <= DL_EPS) OR (fWaterKg <= DL_EPS) OR (fMaltCpKJkgK <= DL_EPS)
   OR (fWaterCpKJkgK <= DL_EPS) OR (fLossPct < DL_ZERO) OR (fLossPct > DL_LOSS_MAX) THEN
    FC_DL_MashStrikeWaterTempCalc := -1.0;  (* 哨兵 -1：组态非法 / Sentinel -1 bad config *)
    RETURN;
END_IF
(* 两侧热容：C = m·cp [kJ/K] *)
fHeatCapMaltKJK  := fMaltKg * fMaltCpKJkgK;
fHeatCapWaterKJK := fWaterKg * fWaterCpKJkgK;
(* 热损修正：需把目标温度按热损率上调，等效为多带入焓 *)
fLossUnit := fLossPct / DL_PCT_BASE;
fTargetEffC := fTargetMashC * (1.0 + fLossUnit);
(* 能量平衡：T_w = [T_eff·(Cm+Cw) - Cm·Tm] / Cw，除子水热容已过域闸 *)
fStrikeWaterC := (fTargetEffC * (fHeatCapMaltKJK + fHeatCapWaterKJK)
                  - fHeatCapMaltKJK * fMaltT0C) / fHeatCapWaterKJK;
xValid := TRUE;                                 (* 链路有效 / Chain valid *)
FC_DL_MashStrikeWaterTempCalc := fStrikeWaterC; (* 返回投料水温 [°C] / Return strike water temp *)
END_FUNCTION

(* ---- FC_DL_MembraneFluxCalc.st ---- *)
(*
  ============================================================
  组件名 : FC_DL_MembraneFluxCalc
  分类   : DL_Process
  功能   : 膜通量计算，由产水流量与膜面积求通量并折算相对基准通量的比值
  开源溯源 : internal-design（本轮无外部代码逐行引用）
             参考语义 : 无外部参考
  复杂度 : C1
  版本   : 1.0.0
  ============================================================
*)

FUNCTION FC_DL_MembraneFluxCalc : REAL
VAR_INPUT
    rPermeateFlow_m3h : REAL; // 产水流量 [m3/h] permeate flow [m3 per hour]
    rMembraneArea_m2  : REAL; // 膜面积 [m2] membrane area [m2]
    rFluxRef          : REAL; // 基准通量 [L/m2/h] reference flux [litre per square metre per hour]
END_VAR
VAR_OUTPUT
    rFluxLmh   : REAL; // 实测通量 [L/m2/h] measured flux [litre per square metre per hour]
    rFluxRatio : REAL; // 通量与基准之比 [无量纲] ratio of the flux to the reference [dimensionless]
    bValid     : BOOL; // 结果有效标志 result validity flag
END_VAR
VAR CONSTANT
    DL_M3_TO_L : REAL := 1000.0; // 每立方米升数 litres per cubic metre
END_VAR
VAR
    _bFin : BOOL := FALSE; // 三输入有限性判定 finiteness verdict of the three inputs
    _rFlux: REAL := 0.0; // 通量中间量 [L/m2/h] intermediate flux [litre per square metre per hour]
    _rRat : REAL := 0.0; // 比值中间量 [无量纲] intermediate ratio [dimensionless]
END_VAR

// 段 1｜出口预置 preset the exit
FC_DL_MembraneFluxCalc := 0.0; // 缺省返回零 default zero return
rFluxLmh := 0.0; // 通量预置零 flux preset to zero
rFluxRatio := 0.0; // 比值预置零 ratio preset to zero
bValid := FALSE; // 计算完成前不认结果 unusable before the calculation
// 段 2｜非有限闸 finiteness gate
_bFin := (rPermeateFlow_m3h = rPermeateFlow_m3h) AND (rMembraneArea_m2 = rMembraneArea_m2) AND (rFluxRef = rFluxRef); // 三输入自反判定 self comparison of the three inputs
IF NOT _bFin THEN
    RETURN; // 非有限即无效 non finite means invalid
END_IF
// 段 3｜面积与流量闸 area and flow gate
IF (rMembraneArea_m2 <= 0.0) OR (rPermeateFlow_m3h < 0.0) THEN
    RETURN; // 面积非正或负流量属配置非法 an illegal area or a negative flow
END_IF
// 段 4｜主体通量 main flux
_rFlux := rPermeateFlow_m3h * DL_M3_TO_L / rMembraneArea_m2; // 流量折算升后除面积 flow in litres over the area
rFluxLmh := _rFlux; // 通量落定 land the flux
// 段 5｜基准比值闸 reference ratio gate
IF rFluxRef <= 0.0 THEN
    RETURN; // 基准通量非正无法求比值 a non positive reference cannot carry a ratio
END_IF
_rRat := _rFlux / rFluxRef; // 实测对基准比值 measured over reference
rFluxRatio := _rRat; // 比值落定 land the ratio
bValid := TRUE; // 结果可用 result usable
FC_DL_MembraneFluxCalc := _rFlux; // 函数返回通量 return the flux
END_FUNCTION

(* ---- FC_DL_MembraneTmpCalc.st ---- *)
(*
  ============================================================
  组件名 : FC_DL_MembraneTmpCalc
  分类   : DL_Process
  功能   : 膜系统跨膜压差计算，进料侧取单点或浓水与进料均值，再扣除渗透压得净推动力
  开源溯源 : internal-design（本轮无外部代码逐行引用）
             参考语义 : 无外部参考
  复杂度 : C1
  版本   : 1.0.0
  ============================================================
*)

FUNCTION FC_DL_MembraneTmpCalc : REAL
VAR_INPUT
    rFeedPress_bar : REAL; // 进料侧压力 [bar] feed side pressure [bar]
    rConcPress_bar : REAL; // 浓水侧压力 [bar] concentrate side pressure [bar]
    rPermPress_bar : REAL; // 产水侧压力 [bar] permeate side pressure [bar]
    rOsmotic_bar   : REAL; // 渗透压 [bar] osmotic pressure [bar]
    bUseAvgFeed    : BOOL; // 真为进料与浓水取均值，假为取进料压力 average the feed and the concentrate when true
END_VAR
VAR_OUTPUT
    rTmp_bar       : REAL; // 跨膜压差 [bar] trans membrane pressure [bar]
    rNetDriving_bar: REAL; // 净推动力 [bar] net driving pressure [bar]
    bValid         : BOOL; // 结果有效标志 result validity flag
END_VAR
VAR CONSTANT
    DL_HALF : REAL := 0.5; // 均值系数 averaging factor
END_VAR
VAR
    _bFin   : BOOL := FALSE; // 四实数输入有限性判定 finiteness verdict of the four real inputs
    _rFeed  : REAL := 0.0; // 进料侧有效压力 [bar] effective feed side pressure [bar]
    _rTmp   : REAL := 0.0; // 跨膜压差中间量 [bar] intermediate trans membrane pressure [bar]
    _rNet   : REAL := 0.0; // 净推动力中间量 [bar] intermediate net driving pressure [bar]
END_VAR

// 段 1｜出口预置 preset the exit
FC_DL_MembraneTmpCalc := 0.0; // 缺省返回零 default zero return
rTmp_bar := 0.0; // 跨膜压差预置零 trans membrane pressure preset to zero
rNetDriving_bar := 0.0; // 净推动力预置零 net driving pressure preset to zero
bValid := FALSE; // 计算完成前不认结果 unusable before the calculation
// 段 2｜非有限闸 finiteness gate
_bFin := (rFeedPress_bar = rFeedPress_bar) AND (rConcPress_bar = rConcPress_bar) AND (rPermPress_bar = rPermPress_bar) AND (rOsmotic_bar = rOsmotic_bar); // 四输入自反判定 self comparison of the four inputs
IF NOT _bFin THEN
    RETURN; // 非有限即无效 non finite means invalid
END_IF
// 段 3｜压力方向闸 pressure direction gate
IF (rFeedPress_bar < 0.0) OR (rConcPress_bar < 0.0) OR (rPermPress_bar < 0.0) OR (rOsmotic_bar < 0.0) THEN
    RETURN; // 负压力或负渗透压属配置非法 a negative pressure or osmotic value is illegal
END_IF
// 段 4｜进料侧有效压力选择 the effective feed side pressure
IF bUseAvgFeed THEN
    _rFeed := (rFeedPress_bar + rConcPress_bar) * DL_HALF; // 进料与浓水取均值 average the feed and the concentrate
ELSE
    _rFeed := rFeedPress_bar; // 直接取进料压力 take the feed pressure itself
END_IF
// 段 5｜跨膜压差与净推动力 trans membrane pressure and the net driving force
_rTmp := _rFeed - rPermPress_bar; // 进料侧减产水侧 feed side minus permeate side
rTmp_bar := _rTmp; // 跨膜压差落定 land the trans membrane pressure
_rNet := _rTmp - rOsmotic_bar; // 扣除渗透压 deduct the osmotic pressure
rNetDriving_bar := _rNet; // 净推动力落定 land the net driving force
IF _rTmp > 0.0 THEN
    bValid := TRUE; // 正跨膜压差判结果可用 a positive pressure makes the result usable
END_IF
FC_DL_MembraneTmpCalc := _rTmp; // 函数返回跨膜压差 return the trans membrane pressure
END_FUNCTION

(* ---- FC_DL_MercerCausticPickupCalc.st ---- *)
(*
  Name: FC_DL_MercerCausticPickupCalc
  Category: DL_Process
  Version: 1.0.0
  Round: R91 / 2026-11-25
  开源溯源：clean-room 自研（族 间歇式溢流染色与丝光整理，ST 开源生态实测 0 命中，无外部代码引入）
  功能：1) 丝光碱液带液量（带碱率）按「轧余率 × 碱浓度 / 碱液密度」计算：
           pickup[g/kg 布] = (fPickupPct / 100) * fConcGpl / fDensityKgl，
           其中 fPickupPct 为轧余率（带液量占布重的百分数）、fConcGpl 为碱质量浓度 [g/L]、
           fDensityKgl 为碱液密度 [kg/L]。
           量纲推导： (kg液/kg布) * (g/L) / (kg/L) = (kg液/kg布) * (g/kg液) = g/kg布，故无额外折算因子。
        2) 派生量：fLiquorKgKg = 每公斤布带走的碱液质量 [kg/kg]，用于核算碱液损耗与回收负荷。
        3) 工艺域判定：带碱率低于 fPickupMinGkg 判丝光不足（纤维膨化不够、光泽与尺寸稳定性差），
           高于 fPickupMaxGkg 判过轧（碱耗高、后续中和负荷大）。
  边界条件：1) 非有限值闸：五路实值入参先过 NOT(x > -DL_BIG AND x < DL_BIG)，同时拦 NaN 与 Inf，
           命中即闸断实值通路（带碱率与带液量强制 0.0 且置不足位，保守侧），不得只置标志（R19）。
        2) 密度零闸：fDensityKgl 必须 > DL_EPS（带碱率式的分母），为零则结果发散，判无效。
        3) 浓度量级闸：fConcGpl 必须落在 (0.0, DL_CONC_HI_GPL) 内 ——
           丝光碱浓工程带约 180 ~ 300 g/L，越域说明单位用错（g/L 与 %(w/w) 混用）或测点失效。
        4) 轧余率域闸：fPickupPct 必须落在 [0.0, DL_PICKUP_HI_PCT] 内（超过 200 % 不具物理意义）。
        5) 工艺域闸：须满足 0.0 < fPickupMinGkg < fPickupMaxGkg，越域判无效（判据重叠则永不同时报）。
        6) 判据取原始值（R24）：工艺域判定使用钳制前的 _fPickupRawGkg，钳制只作用于输出。
  量纲自证：见功能 1) 的量纲推导，最终量纲为 g/kg（每公斤布带的纯碱克数）；
           fLiquorKgKg = (kg 液)/(kg 布) = kg/kg，无因次质量比。
  修订历史 Revision :
    2026-11-25  v1.0.0  R91 首版
*)

FUNCTION FC_DL_MercerCausticPickupCalc : BOOL
VAR_INPUT
    fPickupPct       : REAL;   // 轧余率（带液量占布重百分比）[%] / Wet pickup percentage [%]
    fConcGpl         : REAL;   // 碱液质量浓度 [g/L] / Caustic mass concentration [g/L]
    fDensityKgl      : REAL;   // 碱液密度 [kg/L] / Caustic liquor density [kg/L]
    fPickupMinGkg    : REAL;   // 带碱率工艺下限 [g/kg] / Caustic pickup process low limit [g/kg]
    fPickupMaxGkg    : REAL;   // 带碱率工艺上限 [g/kg] / Caustic pickup process high limit [g/kg]
END_VAR
VAR_OUTPUT
    fPickupGkg       : REAL;   // 带碱率（每公斤布的纯碱克数）[g/kg] / Caustic pickup per kg of fabric [g/kg]
    fLiquorKgKg      : REAL;   // 每公斤布带走的碱液质量 [kg/kg] / Caustic liquor carried per kg of fabric [kg/kg]
    xPickupLow       : BOOL;   // 带碱率不足标志 [bool] / Caustic pickup below the low limit flag [bool]
    xPickupHigh      : BOOL;   // 带碱率过高标志 [bool] / Caustic pickup above the high limit flag [bool]
    xValid           : BOOL;   // 计算有效标志 [bool] / Calculation valid flag [bool]
END_VAR
VAR
    _fLiquorRawKgKg  : REAL;   // 钳制前的带液量 [kg/kg] / Raw liquor mass ratio before limiting [kg/kg]
    _fPickupRawGkg   : REAL;   // 钳制前的带碱率 [g/kg] / Raw caustic pickup before limiting [g/kg]
END_VAR
VAR CONSTANT
    DL_EPS           : REAL := 1.0E-9;    // 数值零闸阈值 [-] / Numeric zero gate threshold [-]
    DL_BIG           : REAL := 1.0E12;    // 非有限值闸量级上限 [-] / Finiteness gate magnitude [-]
    DL_PCT           : REAL := 100.0;     // 百分比换算因子 [%] / Percent conversion factor [%]
    DL_CONC_HI_GPL   : REAL := 1000.0;    // 碱浓量级闸上限 [g/L] / Concentration magnitude upper bound [g/L]
    DL_PICKUP_HI_PCT : REAL := 200.0;     // 轧余率物理上限 [%] / Wet pickup physical upper bound [%]
    DL_PICKUP_HI_GKG : REAL := 1000.0;    // 带碱率物理上限 [g/kg] / Caustic pickup upper bound [g/kg]
END_VAR

(* —— 段 1：非有限值闸（R19：闸断实值通路；失效侧置不足位，保守侧） —— *)
IF NOT (fPickupPct > -DL_BIG AND fPickupPct < DL_BIG)
   OR NOT (fConcGpl > -DL_BIG AND fConcGpl < DL_BIG)
   OR NOT (fDensityKgl > -DL_BIG AND fDensityKgl < DL_BIG)
   OR NOT (fPickupMinGkg > -DL_BIG AND fPickupMinGkg < DL_BIG)
   OR NOT (fPickupMaxGkg > -DL_BIG AND fPickupMaxGkg < DL_BIG) THEN
    fPickupGkg := 0.0;                      // 输出强制 0.0，切断污染源 / Force zero, cut polluted path
    fLiquorKgKg := 0.0;                     // 带液量强制 0.0 / Liquor ratio forced to zero
    xPickupLow := TRUE;                     // 失效侧按不足处理（保守侧）/ Treat as insufficient when invalid
    xPickupHigh := FALSE;                   // 失效侧过高位保持假 / High flag stays false
    xValid := FALSE;                        // 有效位清零 / Validity cleared
    FC_DL_MercerCausticPickupCalc := FALSE; // 返回码与有效位同源 / Return mirrors validity
    RETURN;                                 // 立即退出 / Immediate exit
END_IF

(* —— 段 2：密度零闸与域闸（密度为带碱率分母） —— *)
IF (fDensityKgl <= DL_EPS)                                        // 密度不可为零
   OR (fConcGpl <= 0.0)                                           // 碱浓必须为正（无碱即无丝光）
   OR (fConcGpl > DL_CONC_HI_GPL)                                 // 碱浓不得超量级闸
   OR (fPickupPct < 0.0)                                          // 轧余率不得为负
   OR (fPickupPct > DL_PICKUP_HI_PCT)                             // 轧余率不得超物理上限
   OR (fPickupMinGkg <= 0.0)                                      // 工艺下限必须为正
   OR (fPickupMaxGkg <= fPickupMinGkg) THEN                       // 工艺上限必须严格大于下限
    fPickupGkg := 0.0;                      // 参数不可用即不可算 / No parameter, no pickup
    fLiquorKgKg := 0.0;                     // 带液量不可算 / Liquor ratio not computable
    xPickupLow := TRUE;                     // 按不足处理（保守侧）/ Treat as insufficient
    xPickupHigh := FALSE;                   // 过高位保持假 / High flag stays false
    xValid := FALSE;                        // 判无效 / Invalid
    FC_DL_MercerCausticPickupCalc := FALSE; // 返回码同步 / Return synchronised
    RETURN;                                 // 提前退出 / Early exit
END_IF

(* —— 段 3：主算式（不钳制，先出原始值供段 4 判据使用，R24） —— *)
_fLiquorRawKgKg := fPickupPct / DL_PCT;                                           // 带液量 [kg/kg]
_fPickupRawGkg := _fLiquorRawKgKg * fConcGpl / fDensityKgl;                        // 带碱率 [g/kg]

(* —— 段 4：判据（取原始值；单点 BOOL 聚合避免多处赋 FALSE 覆盖） —— *)
xPickupLow := (_fPickupRawGkg < fPickupMinGkg);                                    // 丝光不足
xPickupHigh := (_fPickupRawGkg > fPickupMaxGkg);                                   // 过轧
xValid := (_fPickupRawGkg >= 0.0)                                                  // 带碱率不得为负
          AND (_fPickupRawGkg <= DL_PICKUP_HI_GKG)                                 // 不超物理上限（量级异常）
          AND (fPickupMaxGkg <= DL_PICKUP_HI_GKG)                                  // 工艺上限须在物理域内
          AND (_fLiquorRawKgKg >= 0.0);                                            // 带液量不得为负

(* —— 段 5：输出单点写盘（钳制到物理域内，判定结果已在段 4 定案） —— *)
fPickupGkg := LIMIT(0.0, _fPickupRawGkg, DL_PICKUP_HI_GKG);                        // 带碱率钳物理域 [g/kg]
fLiquorKgKg := LIMIT(0.0, _fLiquorRawKgKg, DL_PICKUP_HI_PCT / DL_PCT);             // 带液量钳物理域 [kg/kg]
FC_DL_MercerCausticPickupCalc := xValid;                                           // 返回码：TRUE = 计算可信

END_FUNCTION

(* ---- FC_DL_MercerShrinkageCalc.st ---- *)
(*
  Name: FC_DL_MercerShrinkageCalc
  Category: DL_Process
  Version: 1.0.0
  Round: R91 / 2026-11-25
  开源溯源：clean-room 自研（族 间歇式溢流染色与丝光整理，ST 开源生态实测 0 命中，无外部代码引入）
  功能：1) 丝光收缩率按「经纬密度变化」反算：丝光使纤维膨化、纱线屈曲减少，
           单位长度内纱线根数（密度）上升，故收缩率 = (D_after − D_before) / D_after * 100，
           分母取丝光后密度（即按成品基准计），与纺织行业「按成品计收缩」的惯例一致。
        2) 经纬分别输出 fWarpShrinkPct（经向）/ fWeftShrinkPct（纬向），并给出算术平均
           fAvgShrinkPct，供工艺判断丝光均匀性（经纬差过大说明张力控制不一致）。
        3) 负值判异常：密度减少（收缩率为负）在丝光工序物理上不可能（丝光只增密不疏松），
           判 xNegative = TRUE 且 xValid = FALSE，不取绝对值掩盖方向错误。
  边界条件：1) 非有限值闸：四路实值入参先过 NOT(x > -DL_BIG AND x < DL_BIG)，同时拦 NaN 与 Inf，
           命中即闸断实值通路（三个收缩率强制 0.0），不得只置标志（R19）。
        2) 分母零闸：丝光后密度 fWarpDensityAfter / fWeftDensityAfter 均须 > DL_EPS
           （收缩率式的分母），为零则结果发散，判无效。
        3) 密度非负闸：丝光前密度不得为负（负密度属测点或录入错误），判无效。
        4) 判据取原始值（R24）：负值与量级判定使用钳制前的原始收缩率，钳制只作用于输出。
        5) 物理域钳制：收缩率钳 -DL_SHRINK_SPAN ~ +DL_SHRINK_SPAN（±100 %），
           保留负值观测余量以供上层识别异常方向。
        6) 纯函数无状态：多批次收缩率的统计与工艺纠偏由上层质量模块承担。
  量纲自证：shrink = (根/10cm − 根/10cm) / (根/10cm) * 100 = 无因次百分数 [%]，
           比量上下同为密度量纲（纱线根数/10cm），量纲合法。
  修订历史 Revision :
    2026-11-25  v1.0.0  R91 首版
*)

FUNCTION FC_DL_MercerShrinkageCalc : BOOL
VAR_INPUT
    fWarpDensityBefore : REAL;   // 丝光前经密 [ends/10cm] / Warp density before mercerising [ends/10cm]
    fWarpDensityAfter  : REAL;   // 丝光后经密 [ends/10cm] / Warp density after mercerising [ends/10cm]
    fWeftDensityBefore : REAL;   // 丝光前纬密 [picks/10cm] / Weft density before mercerising [picks/10cm]
    fWeftDensityAfter  : REAL;   // 丝光后纬密 [picks/10cm] / Weft density after mercerising [picks/10cm]
END_VAR
VAR_OUTPUT
    fWarpShrinkPct   : REAL;   // 经向收缩率 [%] / Warp shrinkage [%]
    fWeftShrinkPct   : REAL;   // 纬向收缩率 [%] / Weft shrinkage [%]
    fAvgShrinkPct    : REAL;   // 经纬平均收缩率 [%] / Average shrinkage of warp and weft [%]
    xNegative        : BOOL;   // 出现负收缩（方向异常）标志 [bool] / Negative shrinkage flag [bool]
    xValid           : BOOL;   // 计算有效标志 [bool] / Calculation valid flag [bool]
END_VAR
VAR
    _fWarpRawPct     : REAL;   // 钳制前的经向收缩率 [%] / Raw warp shrinkage before limiting [%]
    _fWeftRawPct     : REAL;   // 钳制前的纬向收缩率 [%] / Raw weft shrinkage before limiting [%]
    _fAvgRawPct      : REAL;   // 钳制前的平均收缩率 [%] / Raw average before limiting [%]
END_VAR
VAR CONSTANT
    DL_EPS           : REAL := 1.0E-9;    // 数值零闸阈值 [-] / Numeric zero gate threshold [-]
    DL_BIG           : REAL := 1.0E12;    // 非有限值闸量级上限 [-] / Finiteness gate magnitude [-]
    DL_PCT           : REAL := 100.0;     // 百分比换算因子 [%] / Percent conversion factor [%]
    DL_TWO           : REAL := 2.0;       // 平均值折算系数 [-] / Average divisor [-]
    DL_DENS_HI       : REAL := 5000.0;    // 密度量级闸上限 [ends/10cm] / Density magnitude upper bound [ends/10cm]
    DL_SHRINK_SPAN   : REAL := 100.0;     // 收缩率钳制跨度 [%] / Shrinkage clamp span [%]
END_VAR

(* —— 段 1：非有限值闸（R19：闸断实值通路） —— *)
IF NOT (fWarpDensityBefore > -DL_BIG AND fWarpDensityBefore < DL_BIG)
   OR NOT (fWarpDensityAfter > -DL_BIG AND fWarpDensityAfter < DL_BIG)
   OR NOT (fWeftDensityBefore > -DL_BIG AND fWeftDensityBefore < DL_BIG)
   OR NOT (fWeftDensityAfter > -DL_BIG AND fWeftDensityAfter < DL_BIG) THEN
    fWarpShrinkPct := 0.0;                  // 输出强制 0.0，切断污染源 / Force zero, cut polluted path
    fWeftShrinkPct := 0.0;                  // 纬向强制 0.0 / Weft forced to zero
    fAvgShrinkPct := 0.0;                   // 平均强制 0.0 / Average forced to zero
    xNegative := TRUE;                      // 失效侧按方向异常处理（保守侧）/ Treat as abnormal when invalid
    xValid := FALSE;                        // 有效位清零 / Validity cleared
    FC_DL_MercerShrinkageCalc := FALSE;     // 返回码与有效位同源 / Return mirrors validity
    RETURN;                                 // 立即退出 / Immediate exit
END_IF

(* —— 段 2：分母零闸与量级闸（分母取丝光后密度） —— *)
IF (fWarpDensityAfter <= DL_EPS)                                  // 后经密不可为零
   OR (fWeftDensityAfter <= DL_EPS)                               // 后纬密不可为零
   OR (fWarpDensityBefore < 0.0)                                  // 前经密不得为负
   OR (fWeftDensityBefore < 0.0)                                  // 前纬密不得为负
   OR (fWarpDensityAfter > DL_DENS_HI)                            // 后经密量级闸
   OR (fWeftDensityAfter > DL_DENS_HI)                            // 后纬密量级闸
   OR (fWarpDensityBefore > DL_DENS_HI)                           // 前经密量级闸
   OR (fWeftDensityBefore > DL_DENS_HI) THEN                      // 前纬密量级闸
    fWarpShrinkPct := 0.0;                  // 分母为零即不可算 / No denominator, no ratio
    fWeftShrinkPct := 0.0;                  // 纬向不可算 / Weft not computable
    fAvgShrinkPct := 0.0;                   // 平均不可算 / Average not computable
    xNegative := TRUE;                      // 按方向异常处理（保守侧）/ Treat as abnormal
    xValid := FALSE;                        // 判无效 / Invalid
    FC_DL_MercerShrinkageCalc := FALSE;     // 返回码同步 / Return synchronised
    RETURN;                                 // 提前退出 / Early exit
END_IF

(* —— 段 3：主算式（不钳制，先出原始值供段 4 判据使用，R24） —— *)
_fWarpRawPct := (fWarpDensityAfter - fWarpDensityBefore) / fWarpDensityAfter * DL_PCT;   // 经向 [%]
_fWeftRawPct := (fWeftDensityAfter - fWeftDensityBefore) / fWeftDensityAfter * DL_PCT;   // 纬向 [%]
_fAvgRawPct := (_fWarpRawPct + _fWeftRawPct) / DL_TWO;                                   // 平均 [%]

(* —— 段 4：判据（取原始值；单点 BOOL 聚合避免多处赋 FALSE 覆盖） —— *)
xNegative := (_fWarpRawPct < 0.0) OR (_fWeftRawPct < 0.0);                        // 密度减少：方向异常
xValid := (NOT xNegative)                                                         // 丝光只增密不疏松
          AND (_fWarpRawPct <= DL_SHRINK_SPAN)                                    // 不超钳制跨度（量级异常）
          AND (_fWeftRawPct <= DL_SHRINK_SPAN)                                    // 不超钳制跨度
          AND (_fAvgRawPct >= 0.0);                                               // 平均值非负（与方向闸一致）

(* —— 段 5：输出单点写盘（钳制到物理域内，判定结果已在段 4 定案） —— *)
fWarpShrinkPct := LIMIT(-DL_SHRINK_SPAN, _fWarpRawPct, DL_SHRINK_SPAN);            // 经向钳 ±100 [%]
fWeftShrinkPct := LIMIT(-DL_SHRINK_SPAN, _fWeftRawPct, DL_SHRINK_SPAN);            // 纬向钳 ±100 [%]
fAvgShrinkPct := LIMIT(-DL_SHRINK_SPAN, _fAvgRawPct, DL_SHRINK_SPAN);              // 平均钳 ±100 [%]
FC_DL_MercerShrinkageCalc := xValid;                                              // 返回码：TRUE = 计算可信

END_FUNCTION

(* ---- FC_DL_MethaneRatioCalc.st ---- *)
(*
  道莅工业代码库 / Daoli Industrial ST Library
  组件: FC_DL_MethaneRatioCalc
  分类: DL_Process
  开源溯源: 无（clean-room 工程公式自研；参考公开工艺计算公式，未复制任何受版权保护代码）
  许可证: 本项目自有 (MIT)
  功能: 沼气组分平衡求甲烷含量与低位热值 LHV，含 H2S 腐蚀告警
*)
FUNCTION FC_DL_MethaneRatioCalc : BOOL
VAR_INPUT
    rCo2Pct : REAL; // 二氧化碳体积分数 [%] / CO2 volume fraction
    rN2Pct : REAL; // 氮气体积分数 [%] / N2 volume fraction
    rO2Pct : REAL; // 氧气体积分数 [%] / O2 volume fraction
    rH2sPpm : REAL; // 硫化氢浓度 [ppm] / H2S concentration in ppm
END_VAR
VAR_OUTPUT
    rCh4Pct : REAL; // 甲烷体积分数 [%] / methane volume fraction
    rLhvMJm3 : REAL; // 低位热值 [MJ/m3] / lower heating value
    bValid : BOOL; // 结果有效位 [-] / result valid flag
    iErrCode : INT; // 事件码 0=正常 1=组分和超 100（甲烷按 0 饱和）2=H2S 超 500ppm 告警 3=结果非有限 / event code
END_VAR
VAR CONSTANT
    rPctFull : REAL := 100.0; // 组分满量程 [%] / full scale of volume fraction
    rCh4Lhv : REAL := 35.8; // 纯甲烷低位热值 [MJ/m3] / LHV of pure methane
    rH2sLimit : REAL := 500.0; // H2S 腐蚀告警门槛 [ppm] / H2S corrosion alarm threshold
    rPctToFrac : REAL := 0.01; // 百分数转小数系数 [-]/[%] / percent to fraction factor
END_VAR
VAR
    rSumPct : REAL; // 非甲烷组分之和 [%] / sum of non-methane fractions
    rCh4Raw : REAL; // 未饱和甲烷含量 [%] / unlimited methane fraction
END_VAR

    // —— 段 0：全路径预清 —— //
    rSumPct := 0.0;
    rCh4Raw := 0.0;
    rCh4Pct := 0.0;
    rLhvMJm3 := 0.0;
    bValid := FALSE;
    iErrCode := 0;
    FC_DL_MethaneRatioCalc := FALSE;
    // —— 段 1：量纲链 (% + % + %) = % —— //
    rSumPct := rCo2Pct + rN2Pct + rO2Pct; // 非甲烷组分和 [%] / non-methane sum
    // —— 段 2：组分和非负性与满量程闸 —— //
    IF rSumPct < 0.0 THEN
        iErrCode := 1; // 组分和为负，分析仪故障 / negative sum, analyser fault
        RETURN;
    END_IF;
    rCh4Raw := rPctFull - rSumPct; // 甲烷 = 100 - 其余 [%] / methane by difference
    // —— 段 3：甲烷负值饱和为 0 并置信息码 —— //
    IF (rCo2Pct < 0.0) OR (rN2Pct < 0.0) OR (rO2Pct < 0.0) THEN
        iErrCode := 4; // 组分负值：传感器非法，甲烷不可信 / negative component: invalid sensor
        bValid := FALSE;
        FC_DL_MethaneRatioCalc := TRUE;
        RETURN;
    END_IF
    IF rCh4Raw > 100.0 THEN
        rCh4Pct := 100.0; // 组分和偏低导致外推超 100%，饱和 / extrapolated above 100 percent, clamp
    ELSIF rCh4Raw < 0.0 THEN
        rCh4Pct := 0.0;
        iErrCode := 1; // 组分和超 100%，甲烷按零饱和 / sum above 100 percent, methane floored at zero
    ELSE
        rCh4Pct := rCh4Raw;
    END_IF;
    // —— 段 4：热值 (MJ/m3) = 甲烷份额 × 纯甲烷 LHV；H2S 告警 —— //
    rLhvMJm3 := rCh4Pct * rPctToFrac * rCh4Lhv; // 低位热值 [MJ/m3] / lower heating value
    IF ABS(rLhvMJm3) > 1.0E15 THEN
        rLhvMJm3 := 0.0;
        iErrCode := 3; // 结果非有限，强制归零 / non-finite result, forced to zero
        RETURN;
    END_IF;
    IF rH2sPpm > rH2sLimit THEN
        iErrCode := 2; // 信息级：H2S 超限，注意脱硫与腐蚀 / info: H2S high, check desulfurisation
    END_IF;
    bValid := TRUE;
    FC_DL_MethaneRatioCalc := TRUE;
END_FUNCTION

(* ---- FC_DL_MoldClampForceCalc.st ---- *)
(*
 * FC_DL_MoldClampForceCalc | C2 | DL_Process
 * 功能：浇注时铁水浮力（抬箱力）与合型压铁力（含安全系数）       单位：体积 [L]、密度 [kg/L]、重力 [m/s²]、力 [kN]、安全系数 [1]
 * 工况边界：按等效液柱静压简化 F=V×ρ×g（未计浇口杯高度附加压头与冲击动压）；型腔体积与安全系数须 >0、密度须 >0 且有限；小件压铁力偏小属正常，须由工艺员叠加砂箱自重判定
 * 代数值回代：V=12 L、ρ=7.0 kg/L、g=9.80665 → F=12×7×9.80665/1000=0.824 kN；SF=1.5 → clamp=1.24 kN（与 spec 回代行一致）
 * 开源溯源：clean-room 自研，未复制任何第三方代码（无外部来源）
 *)
FUNCTION FC_DL_MoldClampForceCalc : BOOL
VAR_INPUT
    rCavityVolL      : REAL := 12.0;      // 型腔体积 | mould cavity volume [L]
    rMetalDensityKgL : REAL := 7.0;       // 铁水密度 | molten iron density [kg/L]
    rGravity         : REAL := 9.80665;   // 重力加速度 | gravitational acceleration [m/s²]
    rSf              : REAL := 1.5;       // 安全系数 | safety factor [1]
END_VAR
VAR_OUTPUT
    rBuoyancyKn : REAL;                   // 抬箱力（浮力）| lifting force [kN]
    rClampKn    : REAL;                   // 压铁力 | clamp force [kN]
    xValid      : BOOL;                   // 输出有效 | outputs valid
END_VAR
VAR
    xFinV   : BOOL;                       // 体积有限性 | volume is finite
    xFinRho : BOOL;                       // 密度有限性 | density is finite
    xFinG   : BOOL;                       // 重力有限性 | gravity is finite
    xFinSf  : BOOL;                       // 安全系数有限性 | safety factor is finite
END_VAR
VAR CONSTANT
    DL_MCF_N_TO_KN : REAL := 1000.0;      // 牛转千牛系数 | newtons to kilonewtons factor [N/kN]
END_VAR

// 段1｜非有限闸（R19）
xFinV := (rCavityVolL = rCavityVolL) AND ((rCavityVolL - rCavityVolL) = 0.0);
xFinRho := (rMetalDensityKgL = rMetalDensityKgL) AND ((rMetalDensityKgL - rMetalDensityKgL) = 0.0);
xFinG := (rGravity = rGravity) AND ((rGravity - rGravity) = 0.0);
xFinSf := (rSf = rSf) AND ((rSf - rSf) = 0.0);
IF (NOT xFinV) OR (NOT xFinRho) OR (NOT xFinG) OR (NOT xFinSf) THEN
    rBuoyancyKn := 0.0;                   // 安全值：力 0 | safe value, zero force
    rClampKn := 0.0;
    xValid := FALSE;
    FC_DL_MoldClampForceCalc := FALSE;
    RETURN;
END_IF

// 段2｜域闸：体积、密度、安全系数须为正，重力须 >0
IF (rCavityVolL <= 0.0) OR (rMetalDensityKgL <= 0.0) OR (rGravity <= 0.0) OR (rSf <= 0.0) THEN
    rBuoyancyKn := 0.0;
    rClampKn := 0.0;
    xValid := FALSE;
    FC_DL_MoldClampForceCalc := FALSE;
    RETURN;
END_IF

// 段3｜算法：F = V×ρ×g/1000 kN；clamp = F×SF
rBuoyancyKn := rCavityVolL * rMetalDensityKgL * rGravity / DL_MCF_N_TO_KN;
rClampKn := rBuoyancyKn * rSf;

// 段4｜出口
xValid := TRUE;
FC_DL_MoldClampForceCalc := TRUE;
END_FUNCTION

(* ---- FC_DL_MotorLoadFactorCalc.st ---- *)
(*
  ============================================================
  组件名 : FC_DL_MotorLoadFactorCalc
  分类   : DL_Process
  功能   : 电机负载率计算，由实测有功功率与功率因数求视在功率并折算负载率与过载位
  复杂度 : C1
  版本   : 1.0.0
  作者   : 道莅工业代码库工厂 / R81
  日期   : 2026-11-24
  开源溯源 : clean-room（no upstream）—— 依据公开工程公式自研，未复制任何上游实现
  红线自检 : R1 无GVL/R2 无物理地址/R3 纯IEC/R4 防除零/R5 双语注释
  接口说明 :
      视在功率 = 有功功率 / 功率因数，功率因数不高于 0.1 视为测量不可信，直接判无效。
      负载率 = 有功 / 额定有功 * 100，限幅 0~150；超过 100% 置过载位。
      限幅上限取 150% 而非 100%，是为了在过载时保留可区分的幅值信息。
  ============================================================
*)
FUNCTION FC_DL_MotorLoadFactorCalc : BOOL
VAR_INPUT
    bEnable   : BOOL; // 使能：TRUE 时计算 / Enable: TRUE to compute
    bErr      : BOOL; // 外部故障：TRUE 时立即退出并置结果无效 / External fault: TRUE aborts with invalid result
    rP_kw     : REAL; // 实测有功功率 [kW] / measured active power [kilowatt]
    rPnom_kw  : REAL; // 电机额定有功功率 [kW] / rated active power of the motor [kilowatt]
    rCosPhi   : REAL; // 实测功率因数 [无量纲] / measured power factor [dimensionless]
END_VAR
VAR_OUTPUT
    rApparentKva : REAL; // 视在功率 [kVA] / apparent power [kilovolt ampere]
    rLoadPct     : REAL; // 负载率，限幅 0~150 [%] / load factor clamped to 0 to 150 [percent]
    bOverload    : BOOL; // 过载：TRUE 表示负载率超过 100% / overload, TRUE when the load factor exceeds 100 percent
    bValid       : BOOL; // 输出有效：TRUE 表示结果可用 / Output valid
END_VAR
VAR CONSTANT
    DL_R_MAX     : REAL := 3.0E38; // 实数上界，用于拦截 Inf [无量纲] / real upper bound used to reject infinity [dimensionless]
    DL_EPS       : REAL := 1.0E-12; // 除零判定阈值 [无量纲] / division guard threshold [dimensionless]
    DL_PF_MIN    : REAL := 0.1;    // 功率因数可信下界 [无量纲] / credible lower bound of the power factor [dimensionless]
    DL_PF_MAX    : REAL := 1.0;    // 功率因数物理上界 [无量纲] / physical upper bound of the power factor [dimensionless]
    DL_PCT       : REAL := 100.0;  // 百分数换算系数 [无量纲] / percentage scaling factor [dimensionless]
    DL_LOAD_HI   : REAL := 150.0;  // 负载率限幅上限 [%] / upper clamp of the load factor [percent]
    DL_LOAD_LO   : REAL := 0.0;    // 负载率限幅下限 [%] / lower clamp of the load factor [percent]
    DL_OVL_PCT   : REAL := 100.0;  // 过载门限 [%] / overload threshold [percent]
END_VAR
VAR
    _bFin  : BOOL := FALSE; // 输入有限性判定结果 / input finiteness verdict
    _rRaw  : REAL := 0.0;   // 限幅前负载率 [%] / raw load factor before clamping [percent]
END_VAR

    // 段 1｜出口预置
    rApparentKva := 0.0;
    rLoadPct := 0.0;
    bOverload := FALSE;
    bValid := FALSE;
    // 段 2｜使能闸与外部故障闸
    IF NOT bEnable THEN
        RETURN;
    END_IF;
    IF bErr THEN
        RETURN;
    END_IF;
    // 段 3｜非有限闸
    _bFin := (rP_kw = rP_kw) AND (ABS(rP_kw) <= DL_R_MAX) AND (rPnom_kw = rPnom_kw) AND (ABS(rPnom_kw) <= DL_R_MAX) AND (rCosPhi = rCosPhi) AND (ABS(rCosPhi) <= DL_R_MAX);
    IF NOT _bFin THEN
        RETURN;
    END_IF;
    // 段 4｜域闸：额定功率严格为正，有功功率非负，功率因数在可信区间
    IF (ABS(rPnom_kw) <= DL_EPS) OR (rPnom_kw < 0.0) THEN
        RETURN;
    END_IF;
    IF rP_kw < 0.0 THEN
        RETURN;
    END_IF;
    IF (rCosPhi <= DL_PF_MIN) OR (rCosPhi > DL_PF_MAX) THEN
        RETURN;
    END_IF;
    // 段 5｜视在功率
    rApparentKva := rP_kw / rCosPhi;
    // 段 6｜负载率与限幅
    _rRaw := rP_kw / rPnom_kw * DL_PCT;
    IF _rRaw < DL_LOAD_LO THEN
        rLoadPct := DL_LOAD_LO;
    ELSIF _rRaw > DL_LOAD_HI THEN
        rLoadPct := DL_LOAD_HI;
    ELSE
        rLoadPct := _rRaw;
    END_IF;
    // 段 7｜过载位用限幅前的真实值判定，避免限幅把过载信息吃掉
    IF _rRaw > DL_OVL_PCT THEN
        bOverload := TRUE;
    ELSE
        bOverload := FALSE;
    END_IF;
    bValid := TRUE;
    FC_DL_MotorLoadFactorCalc := bValid;
END_FUNCTION

(* ---- FC_DL_MtsrCalc.st ---- *)
(*
  DL Factory R84 | FC_DL_MtsrCalc
  功能：由当前温度与绝热温升算 MTSR，并给分解起始温度的安全裕度
  开源溯源：无（clean-room 自研，依据公开工艺公式，来源=行业通用公式，许可证=MIT，借鉴点=公式结构）
  规则：R1-R16 全遵守
*)
FUNCTION FC_DL_MtsrCalc : REAL
VAR_INPUT
    fTpC : REAL := 80.0; // 当前工艺温度 [℃] / current process temperature [C]
    fDTadK : REAL := 60.0; // 绝热温升（由绝热温升计算件给出） [K] / adiabatic temperature rise [K]
    fConvertFrac : REAL := 0.6; // 已转化分数（0~1） [-] / converted fraction [0,1]
    fStartDecompC : REAL := 180.0; // 分解起始温度 [℃] / decomposition onset temperature [C]
    fMarginMinK : REAL := 20.0; // 最小安全裕度门限 [K] / minimum safety margin [K]
END_VAR
VAR_OUTPUT
    fMarginK : REAL; // 安全裕度（分解起始 − MTSR） [K] / safety margin [K]
    xRisk : BOOL; // 裕度不足风险位 [-] / insufficient margin risk flag [-]
    xValid : BOOL; // 计算结果有效标志 [-] / calculation valid flag [-]
END_VAR
VAR
    fUnconvFrac : REAL; // 未转化分数（1 − X，钳位） [-] / unconverted fraction [-]
    fMtsrC : REAL; // MTSR 中间量 [℃] / MTSR intermediate [C]
END_VAR

// 段 1｜出口预置（R256）
FC_DL_MtsrCalc := -1.0; // 哨兵返回 -1（无效） [-] / sentinel return -1, invalid [-]
fMarginK := 0.0; // 裕度预置零 [K] / margin preset zero [K]
xRisk := FALSE; // 风险位预置 FALSE [-] / risk preset false [-]
xValid := FALSE; // 计算完成前不认结果 [-] / unusable before calculation [-]

// 段 2｜非有限拦截 + 域闸（R4/R20）
IF NOT (fTpC > -1.0E30 AND fTpC < 1.0E30) OR NOT (fDTadK > -1.0E30 AND fDTadK < 1.0E30) OR NOT (fConvertFrac > -1.0E30 AND fConvertFrac < 1.0E30) OR NOT (fStartDecompC > -1.0E30 AND fStartDecompC < 1.0E30) OR NOT (fMarginMinK > -1.0E30 AND fMarginMinK < 1.0E30) THEN
    RETURN; // 任一入参为 NaN/Inf 一律拒绝 [-] / any NaN or Inf input rejected [-]
END_IF
IF fDTadK < 0.0 OR fMarginMinK < 0.0 THEN
    RETURN; // 绝热温升与裕度门限非负域闸 [K] / non negative rise and margin gate [K]
END_IF

// 段 3｜未转化分数（钳位 0~1）
fUnconvFrac := 1.0 - fConvertFrac; // 无量纲：1 − [-] = - / dimensionless one minus the fraction
IF fUnconvFrac < 0.0 THEN
    fUnconvFrac := 0.0; // 转化分数超一钳零（无剩余潜热） [-] / clamp low: no residual potential [-]
END_IF
IF fUnconvFrac > 1.0 THEN
    fUnconvFrac := 1.0; // 负转化分数钳一（按全未转化计，保守） [-] / clamp high: assume full potential [-]
END_IF

// 段 4｜MTSR = Tp + ΔTad × (1 − X)
fMtsrC := fTpC + (fDTadK * fUnconvFrac); // ℃ + K × 无量纲 = ℃（温差按同刻度计） / [C] + [K] × [-] = [C]
IF NOT (fMtsrC > -1.0E30 AND fMtsrC < 1.0E30) THEN
    RETURN; // 结果非有限再拦一次 [-] / second finiteness gate [-]
END_IF

// 段 5｜安全裕度与风险位
fMarginK := fStartDecompC - fMtsrC; // ℃ − ℃ = K（温差） / [C] minus [C] = [K]
xRisk := fMarginK < fMarginMinK; // 直比门限，禁浮点等值 [-] / direct compare, no float equality [-]
xValid := TRUE; // 链路有效 [-] / chain valid [-]
FC_DL_MtsrCalc := fMtsrC; // 返回 MTSR [℃] / return the MTSR [C]
END_FUNCTION

(* ---- FC_DL_MullerBatchWeightCalc.st ---- *)
(*
 * FC_DL_MullerBatchWeightCalc | C2 | DL_Process
 * 功能：混砂机单批配比（批量、新砂、膨润土、水、旧砂）       单位：质量 [kg]、比例 [%]、充填系数 [1]
 * 工况边界：单批料量 = 容量×充填系数，充填系数须在 (0,1]；各比例均按「批量」为基数（与 spec 回代一致，水计入批内），三者之和须 ≤100 %，否则判 9712；容量须 >0 且有限
 * 代数值回代：cap=2000 kg、fill=0.75 → batch=1500 kg；新砂 10 %→150 kg；膨润土 1.2 %→18 kg；水 2.8 %→42 kg；旧砂=1500−150−18−42=1290 kg（与 spec 回代行一致）
 * 开源溯源：clean-room 自研，未复制任何第三方代码（无外部来源）
 *)
FUNCTION FC_DL_MullerBatchWeightCalc : BOOL
VAR_INPUT
    rCapacityKg    : REAL := 2000.0;  // 混砂机额定容量 | muller rated capacity [kg]
    rFillFactor    : REAL := 0.75;    // 充填系数 | fill factor [1]
    rNewSandPct    : REAL := 10.0;    // 新砂比例 | new sand ratio [%]
    rBentonitePct  : REAL := 1.2;     // 膨润土比例 | bentonite ratio [%]
    rWaterPct      : REAL := 2.8;     // 水比例 | water ratio [%]
END_VAR
VAR_OUTPUT
    rBatchKg      : REAL;             // 单批料量 | batch weight [kg]
    rNewSandKg    : REAL;             // 新砂加入量 | new sand weight [kg]
    rBentoniteKg  : REAL;             // 膨润土加入量 | bentonite weight [kg]
    rWaterKg      : REAL;             // 水加入量 | water weight [kg]
    rReturnSandKg : REAL;             // 旧砂（回用砂）量 | return sand weight [kg]
    rSumPct       : REAL;             // 三辅料比例之和 | sum of the three additive ratios [%]
    xValid        : BOOL;             // 输出有效 | outputs valid
    nFaultCode    : INT;              // 0=无 / 9712=容量或比例非法 | 0 none, 9712 illegal capacity or ratio
END_VAR
VAR
    xFinCap  : BOOL;                  // 容量有限性 | capacity is finite
    xFinFill : BOOL;                  // 充填系数有限性 | fill factor is finite
    xFinNew  : BOOL;                  // 新砂比例有限性 | new sand ratio is finite
    xFinBent : BOOL;                  // 膨润土比例有限性 | bentonite ratio is finite
    xFinWtr  : BOOL;                  // 水比例有限性 | water ratio is finite
END_VAR
VAR CONSTANT
    DL_MBW_PCT : REAL := 100.0;       // 百分数换算系数 | percentage factor [%]
    DL_MBW_EPS : REAL := 1.0E-6;      // 浮点比较容差 | floating comparison tolerance [%]
END_VAR

// 段1｜非有限闸（R19）
xFinCap := (rCapacityKg = rCapacityKg) AND ((rCapacityKg - rCapacityKg) = 0.0);
xFinFill := (rFillFactor = rFillFactor) AND ((rFillFactor - rFillFactor) = 0.0);
xFinNew := (rNewSandPct = rNewSandPct) AND ((rNewSandPct - rNewSandPct) = 0.0);
xFinBent := (rBentonitePct = rBentonitePct) AND ((rBentonitePct - rBentonitePct) = 0.0);
xFinWtr := (rWaterPct = rWaterPct) AND ((rWaterPct - rWaterPct) = 0.0);
IF (NOT xFinCap) OR (NOT xFinFill) OR (NOT xFinNew) OR (NOT xFinBent) OR (NOT xFinWtr) THEN
    rBatchKg := 0.0;                  // 安全值：全部 0（不配料）| safe value, no batching
    rNewSandKg := 0.0;
    rBentoniteKg := 0.0;
    rWaterKg := 0.0;
    rReturnSandKg := 0.0;
    rSumPct := 0.0;
    xValid := FALSE;
    nFaultCode := 9712;
    FC_DL_MullerBatchWeightCalc := FALSE;
    RETURN;
END_IF

// 段2｜域闸：容量 >0、充填系数 (0,1]、各比例非负且之和 ≤100 %
rSumPct := rNewSandPct + rBentonitePct + rWaterPct;
IF (rCapacityKg <= 0.0) OR (rFillFactor <= 0.0) OR (rFillFactor > 1.0)
   OR (rNewSandPct < 0.0) OR (rBentonitePct < 0.0) OR (rWaterPct < 0.0)
   OR (rSumPct > (DL_MBW_PCT + DL_MBW_EPS)) THEN
    rBatchKg := 0.0;
    rNewSandKg := 0.0;
    rBentoniteKg := 0.0;
    rWaterKg := 0.0;
    rReturnSandKg := 0.0;
    xValid := FALSE;
    nFaultCode := 9712;
    FC_DL_MullerBatchWeightCalc := FALSE;
    RETURN;
END_IF

// 段3｜算法：batch = cap×fill；各辅料按批量比例；旧砂 = 批量 − 三辅料
rBatchKg := rCapacityKg * rFillFactor;
rNewSandKg := rBatchKg * rNewSandPct / DL_MBW_PCT;
rBentoniteKg := rBatchKg * rBentonitePct / DL_MBW_PCT;
rWaterKg := rBatchKg * rWaterPct / DL_MBW_PCT;
rReturnSandKg := rBatchKg - rNewSandKg - rBentoniteKg - rWaterKg;
IF rReturnSandKg < 0.0 THEN
    rReturnSandKg := 0.0;             // 保险钳位（段2的比例和约束已排除）| defensive clamp already excluded by segment 2
END_IF

// 段4｜出口
nFaultCode := 0;
xValid := TRUE;
FC_DL_MullerBatchWeightCalc := TRUE;
END_FUNCTION

(* ---- FC_DL_NozzleClogIndexCalc.st ---- *)
(*
  ============================================================
  组件名 : FC_DL_NozzleClogIndexCalc
  分类   : DL_Process
  功能   : 喷嘴堵塞指数计算，由额定与实测流量求流量偏差率并折算堵塞百分比与报警位
  复杂度 : C1
  版本   : 1.0.0
  作者   : 道莅工业代码库工厂 / R81
  日期   : 2026-11-24
  开源溯源 : clean-room（no upstream）—— 依据公开工程公式自研，未复制任何上游实现
  红线自检 : R1 无GVL/R2 无物理地址/R3 纯IEC/R4 防除零/R5 双语注释
  接口说明 :
      偏差率 = (额定流量 - 实测流量) / 额定流量 * 100，限幅 0~100。
      实测高于额定时偏差为负，属超流而非堵塞，按 0 截断，堵塞指数不会为负。
      堵塞报警门限 15%，严格大于才置位。喷嘴数量仅用于产线级统计，不参与单嘴指数。
  ============================================================
*)
FUNCTION FC_DL_NozzleClogIndexCalc : BOOL
VAR_INPUT
    bEnable     : BOOL; // 使能：TRUE 时计算 / Enable: TRUE to compute
    bErr        : BOOL; // 外部故障：TRUE 时立即退出并置结果无效 / External fault: TRUE aborts with invalid result
    rFlowNom    : REAL; // 额定流量 [L/min] / rated flow [litre per minute]
    rFlowAct    : REAL; // 实测流量 [L/min] / measured flow [litre per minute]
    iNozzleCnt  : INT;  // 参与统计的喷嘴数量 [个] / number of nozzles in the survey [unit]
END_VAR
VAR_OUTPUT
    rDevPct    : REAL; // 限幅前的流量偏差率 [%] / raw flow deviation rate before clamping [percent]
    rClogPct   : REAL; // 堵塞指数，限幅 0~100 [%] / clogging index clamped to 0 to 100 [percent]
    bClogAlarm : BOOL; // 堵塞报警：TRUE 表示指数超过 15% / clog alarm, TRUE when the index exceeds 15 percent
    bValid     : BOOL; // 输出有效：TRUE 表示结果可用 / Output valid
END_VAR
VAR CONSTANT
    DL_R_MAX   : REAL := 3.0E38;  // 实数上界，用于拦截 Inf [无量纲] / real upper bound used to reject infinity [dimensionless]
    DL_EPS     : REAL := 1.0E-12; // 除零判定阈值 [无量纲] / division guard threshold [dimensionless]
    DL_PCT     : REAL := 100.0;   // 百分数换算系数 [无量纲] / percentage scaling factor [dimensionless]
    DL_ZERO    : REAL := 0.0;     // 零值常量 [无量纲] / zero constant [dimensionless]
    DL_ALARM_PCT : REAL := 15.0;  // 堵塞报警门限 [%] / clog alarm threshold [percent]
    DL_MAX_NOZ : INT := 512;      // 喷嘴数量合理上限 [个] / sanity upper bound of the nozzle count [unit]
END_VAR
VAR
    _bFin : BOOL := FALSE; // 输入有限性判定结果 / input finiteness verdict
END_VAR

    // 段 1｜出口预置
    rDevPct := 0.0;
    rClogPct := 0.0;
    bClogAlarm := FALSE;
    bValid := FALSE;
    // 段 2｜使能闸与外部故障闸
    IF NOT bEnable THEN
        RETURN;
    END_IF;
    IF bErr THEN
        RETURN;
    END_IF;
    // 段 3｜非有限闸
    _bFin := (rFlowNom = rFlowNom) AND (ABS(rFlowNom) <= DL_R_MAX) AND (rFlowAct = rFlowAct) AND (ABS(rFlowAct) <= DL_R_MAX);
    IF NOT _bFin THEN
        RETURN;
    END_IF;
    // 段 4｜域闸：额定流量严格为正，实测流量非负，喷嘴数量 1~512
    IF ABS(rFlowNom) <= DL_EPS THEN
        RETURN;
    END_IF;
    IF (rFlowNom < DL_ZERO) OR (rFlowAct < DL_ZERO) THEN
        RETURN;
    END_IF;
    IF (iNozzleCnt < 1) OR (iNozzleCnt > DL_MAX_NOZ) THEN
        RETURN;
    END_IF;
    // 段 5｜偏差率
    rDevPct := (rFlowNom - rFlowAct) / rFlowNom * DL_PCT;
    // 段 6｜限幅到 0~100
    IF rDevPct < DL_ZERO THEN
        rClogPct := DL_ZERO;
    ELSIF rDevPct > DL_PCT THEN
        rClogPct := DL_PCT;
    ELSE
        rClogPct := rDevPct;
    END_IF;
    // 段 7｜报警位
    IF rClogPct > DL_ALARM_PCT THEN
        bClogAlarm := TRUE;
    ELSE
        bClogAlarm := FALSE;
    END_IF;
    bValid := TRUE;
    FC_DL_NozzleClogIndexCalc := bValid;
END_FUNCTION

(* ---- FC_DL_NtuCoagDoseAdj.st ---- *)
(*
  道莅工业代码库 / Daoli Industrial ST Library
  组件: FC_DL_NtuCoagDoseAdj
  分类: DL_Process
  开源溯源: 无（clean-room 工程公式自研；参考公开工艺计算公式，未复制任何受版权保护代码）
  许可证: 本项目自有 (MIT)
  功能: 沉后浊度偏差比例微调混凝投加基准，单次步长与总量双限幅
*)
FUNCTION FC_DL_NtuCoagDoseAdj : BOOL
VAR_INPUT
    rNtuOut : REAL; // 沉后实测浊度 [NTU] / measured settled water turbidity
    rNtuSp : REAL; // 沉后浊度设定值 [NTU] / turbidity setpoint
    rDoseBase : REAL; // 前馈投加基准 [L/h] / feed-forward base dose
    rKp : REAL; // 比例增益 [(L/h)/NTU] / proportional gain
    rStepMax : REAL; // 单次修正步长上限 [L/h] / maximum single-step correction
END_VAR
VAR_OUTPUT
    rDoseOut : REAL; // 修正后投加量 [L/h] / corrected dose
    bValid : BOOL; // 结果有效位 [-] / result valid flag
    iErrCode : INT; // 事件码 0=正常 1=步长上限非法 2=基准投加为负 3=结果非有限 / event code
END_VAR
VAR
    rErr : REAL; // 浊度偏差 实测-设定 [NTU] / turbidity error
    rDelta : REAL; // 比例修正量 [L/h] / proportional correction
    rDoseRaw : REAL; // 未限幅投加量 [L/h] / unlimited dose
    rDoseHi : REAL; // 总量上限 = 2×基准 [L/h] / total upper limit, twice the base
END_VAR

    // —— 段 0：全路径预清 —— //
    rErr := 0.0;
    rDelta := 0.0;
    rDoseRaw := 0.0;
    rDoseHi := 0.0;
    rDoseOut := 0.0;
    bValid := FALSE;
    iErrCode := 0;
    FC_DL_NtuCoagDoseAdj := FALSE;
    // —— 段 1：步长上限闸（限幅基准不可为零） —— //
    IF rStepMax <= 0.0 THEN
        iErrCode := 1; // 步长上限非法，无法限幅 / invalid step limit, clamping impossible
        RETURN;
    END_IF;
    // —— 段 2：基准投加合法性（负基准无物理意义） —— //
    IF rDoseBase < 0.0 THEN
        iErrCode := 2; // 基准投加为负，拒绝修正 / negative base dose rejected
        RETURN;
    END_IF;
    // —— 段 3：比例修正与步长限幅（量纲 (L/h)/NTU × NTU = L/h） —— //
    rErr := rNtuOut - rNtuSp; // 偏差 [NTU] / error
    rDelta := rKp * rErr; // 比例修正 [L/h] / proportional term
    IF rDelta > rStepMax THEN
        rDelta := rStepMax; // 正向步长饱和 / saturate positive step
    ELSIF rDelta < -rStepMax THEN
        rDelta := -rStepMax; // 负向步长饱和 / saturate negative step
    END_IF;
    rDoseRaw := rDoseBase + rDelta; // 修正后投加 [L/h] / corrected dose
    // —— 段 4：总量双限幅 [0, 2×基准] 与结果域闸 —— //
    rDoseHi := rDoseBase + rDoseBase; // 总量上限 [L/h] / total upper limit
    IF ABS(rDoseRaw) > 1.0E15 THEN
        iErrCode := 3; // 结果非有限，强制归零 / non-finite result, forced to zero
        RETURN;
    END_IF;
    IF rDoseRaw < 0.0 THEN
        rDoseOut := 0.0; // 下限零 / floor at zero
    ELSIF rDoseRaw > rDoseHi THEN
        rDoseOut := rDoseHi; // 上限 2×基准 / ceiling at twice the base
    ELSE
        rDoseOut := rDoseRaw;
    END_IF;
    bValid := TRUE;
    FC_DL_NtuCoagDoseAdj := TRUE;
END_FUNCTION

(* ---- FC_DL_OrganicLoadRate.st ---- *)
(*
  道莅工业代码库 / Daoli Industrial ST Library
  组件: FC_DL_OrganicLoadRate
  分类: DL_Process
  开源溯源: 无（clean-room 工程公式自研；参考公开工艺计算公式，未复制任何受版权保护代码）
  许可证: 本项目自有 (MIT)
  功能: 厌氧反应器有机负荷率 OLR（kgVS/(m3·d)）与进料 VS 量计算，含过载判定
*)
FUNCTION FC_DL_OrganicLoadRate : BOOL
VAR_INPUT
    rFeedM3Day : REAL; // 进料体积流量 [m3/d] / feed flow per day
    rCodMgL : REAL; // 进料 COD 浓度 [mg/L] / feed COD concentration
    rVsTsRatio : REAL; // VS/TS 比 [-]，典型 0.7 / volatile to total solids ratio
    rTsKgM3 : REAL; // 进料总固体浓度 [kg/m3] / feed total solids concentration
    rReactorM3 : REAL; // 反应器有效容积 [m3] / reactor working volume
END_VAR
VAR_OUTPUT
    rOlrKgVsM3d : REAL; // 有机负荷率 [kgVS/(m3·d)] / organic loading rate
    rVsKgDay : REAL; // 进料挥发性固体量 [kgVS/d] / volatile solids fed per day
    bValid : BOOL; // 结果有效位 [-] / result valid flag
    bOver : BOOL; // 过载标志（>5.0 kgVS/(m3·d)）[-] / overload flag
    iErrCode : INT; // 事件码 0=正常 1=反应器容积非法 2=VS/TS 比超域 3=结果非有限 / event code
END_VAR
VAR CONSTANT
    rMgLToKgM3 : REAL := 0.001; // mg/L(=g/m3)转 kg/m3 系数 [kg/g] / mg per litre to kg per cubic metre
    rOlrHi : REAL := 5.0; // 过载门槛 [kgVS/(m3·d)] / overload threshold
END_VAR
VAR
    rCodKgM3 : REAL; // 进料 COD 浓度 [kg/m3] / COD concentration in kg/m3
    rVsRaw : REAL; // 未校验 VS 量 [kgVS/d] / unchecked volatile solids
    rOlrRaw : REAL; // 未校验负荷率 [kgVS/(m3·d)] / unchecked loading rate
END_VAR

    // —— 段 0：全路径预清 —— //
    rCodKgM3 := 0.0;
    rVsRaw := 0.0;
    rOlrRaw := 0.0;
    rOlrKgVsM3d := 0.0;
    rVsKgDay := 0.0;
    bValid := FALSE;
    bOver := FALSE;
    iErrCode := 0;
    FC_DL_OrganicLoadRate := FALSE;
    // —— 段 1：分母闸（反应器容积）与 VS/TS 比域闸 —— //
    IF rReactorM3 <= 0.0 THEN
        iErrCode := 1; // 反应器容积非法，负荷率无定义 / invalid reactor volume
        RETURN;
    END_IF;
    IF (rVsTsRatio <= 0.0) OR (rVsTsRatio > 1.0) THEN
        iErrCode := 2; // VS/TS 比超域 (0,1] / VS to TS ratio out of domain
        RETURN;
    END_IF;
    // —— 段 2：量纲链 (m3/d)×(kg/m3)×(-) = kg/d —— //
    rCodKgM3 := rCodMgL * rMgLToKgM3; // COD 浓度 [kg/m3]，仅作参考量 / COD reference only
    // 量纲: (m3/d)*(kg/m3)*(-) = kgVS/d；VS 必须由 TS 乘 VS/TS 得，不得用 COD 冒充
    rVsRaw := rFeedM3Day * rTsKgM3 * rVsTsRatio; // VS 量 [kgVS/d] / volatile solids per day
    IF ABS(rVsRaw) > 1.0E15 THEN
        iErrCode := 3; // 结果非有限，强制归零 / non-finite result, forced to zero
        RETURN;
    END_IF;
    IF rVsRaw < 0.0 THEN
        rVsKgDay := 0.0; // 负进料防御 / negative feed guard
    ELSE
        rVsKgDay := rVsRaw;
    END_IF;
    // —— 段 3：负荷率（量纲 (kg/d)/(m3) = kg/(m3·d)） —— //
    rOlrRaw := rVsKgDay / rReactorM3; // 负荷率 [kgVS/(m3·d)] / organic loading rate
    IF ABS(rOlrRaw) > 1.0E15 THEN
        iErrCode := 3; // 结果非有限，强制归零 / non-finite result, forced to zero
        RETURN;
    END_IF;
    rOlrKgVsM3d := rOlrRaw;
    // —— 段 4：过载判定 —— //
    bOver := rOlrKgVsM3d > rOlrHi; // 过载标志 [-] / overload flag
    bValid := TRUE;
    FC_DL_OrganicLoadRate := TRUE;
END_FUNCTION

(* ---- FC_DL_OverflowDyeFlowCalc.st ---- *)
(*
  Name: FC_DL_OverflowDyeFlowCalc
  Category: DL_Process
  Version: 1.0.0
  Round: R91 / 2026-11-25
  开源溯源：clean-room 自研（族 间歇式溢流染色与丝光整理，ST 开源生态实测 0 命中，无外部代码引入）
  功能：1) 溢流循环流量按喷嘴孔口出流式计算：
           Q = n * Cd * A * SQRT(2 * dP / rho)，
           其中 n 为喷嘴数、Cd 为流量系数（0.6 ~ 0.95）、A 为单孔面积、dP 为泵压折绝对压差 [Pa]、
           rho 为染液密度 [kg/m3]；结果由 m3/s 折算为 m3/h（× 3600）。
           单孔面积由孔径换算：A = pi/4 * d^2，d 以 mm 给出，故需乘 1E-6 折算为 m2。
        2) 派生量：等效喷嘴出口流速 fVelMs 与总开孔面积 fNozzleAreaMm2，
           后者用于判断喷嘴堵塞（面积应与设计值一致，实际流量偏低即堵塞）。
        3) 流量上限保护：结果超过 fFlowMaxM3h 只置 xFlowOver 并钳到上限，
           识别「泵压过高导致超流量」的工况（超流量会拉断布卷并损伤织物组织）。
  边界条件：1) 非有限值闸：四路实值入参先过 NOT(x > -DL_BIG AND x < DL_BIG)，同时拦 NaN 与 Inf，
           命中即闸断实值通路（流量与流速强制 0.0），不得只置标志（R19）。
        2) 孔径零闸：fNozzleDiaMm 必须 > DL_EPS（面积为孔径平方的乘子），
           为零会把「未组态孔径」伪装成「零流量」，判无效而非输出 0。
        3) 密度零闸：fDensityKgm3 必须 > DL_EPS（压差式分母），否则根号内发散。
        4) 系数与数量闸：fDischCoef 必须落在 (0.0, 1.0] 内（大于 1 违反能量守恒）；
           喷嘴数 nNozzle 必须 >= 1（为零即无通路）。
        5) 压差非负闸：fPumpPressKpa 不得为负（负压差会使根号内为负、结果为 NaN），判无效。
        6) 判据取原始值（R24）：超上限判定使用钳制前的 _fFlowRawM3h，钳制只作用于输出。
  量纲自证：A = (mm)^2 * 1E-6 = m2；2*dP/rho = (Pa)/(kg/m3) = (N/m2)*(m3/kg) = m2/s2，
           开方得 m/s；A * v = m2 * m/s = m3/s；再乘 3600 得 m3/h，量纲链闭合。
  修订历史 Revision :
    2026-11-25  v1.0.0  R91 首版
*)

FUNCTION FC_DL_OverflowDyeFlowCalc : BOOL
VAR_INPUT
    nNozzle          : INT;    // 溢流喷嘴数量 [count] / Number of overflow nozzles [count]
    fNozzleDiaMm     : REAL;   // 单喷嘴孔径 [mm] / Single nozzle bore diameter [mm]
    fPumpPressKpa    : REAL;   // 循环泵出口压力（表压）[kPa] / Circulation pump discharge pressure [kPa]
    fDensityKgm3     : REAL;   // 染液密度 [kg/m3] / Dye liquor density [kg/m3]
    fDischCoef       : REAL;   // 喷嘴流量系数（0~1 无因次）[-] / Nozzle discharge coefficient [-]
    fFlowMaxM3h      : REAL;   // 允许循环流量上限 [m3/h] / Permitted circulation flow upper limit [m3/h]
END_VAR
VAR_OUTPUT
    fFlowM3h         : REAL;   // 溢流循环总流量 [m3/h] / Total overflow circulation flow [m3/h]
    fVelMs           : REAL;   // 喷嘴等效出口流速 [m/s] / Equivalent nozzle exit velocity [m/s]
    fNozzleAreaMm2   : REAL;   // 喷嘴总开孔面积 [mm2] / Total nozzle open area [mm2]
    xFlowOver        : BOOL;   // 流量超上限标志 [bool] / Flow overrun flag [bool]
    xValid           : BOOL;   // 计算有效标志 [bool] / Calculation valid flag [bool]
END_VAR
VAR
    _fAreaOneM2      : REAL;   // 单孔面积 [m2] / Single nozzle area [m2]
    _fAreaTotalM2    : REAL;   // 总开孔面积 [m2] / Total open area [m2]
    _fPressPa        : REAL;   // 泵压折算为帕 [Pa] / Pump pressure converted to pascals [Pa]
    _fVelRawMs       : REAL;   // 钳制前的出口流速 [m/s] / Raw exit velocity [m/s]
    _fFlowRawM3s     : REAL;   // 未折算的流量 [m3/s] / Flow before hourly conversion [m3/s]
    _fFlowRawM3h     : REAL;   // 钳制前的原始流量 [m3/h] / Raw flow before limiting [m3/h]
END_VAR
VAR CONSTANT
    DL_EPS           : REAL := 1.0E-9;    // 数值零闸阈值 [-] / Numeric zero gate threshold [-]
    DL_BIG           : REAL := 1.0E12;    // 非有限值闸量级上限 [-] / Finiteness gate magnitude [-]
    DL_PI            : REAL := 3.14159265; // 圆周率 [-] / Pi [-]
    DL_QUARTER       : REAL := 0.25;      // 圆面积折算系数（pi/4 的 1/4 部分）[-] / Circle area factor [-]
    DL_MM2_PER_M2    : REAL := 1.0E6;     // 平方米到平方毫米的折算 [mm2/m2] / Square mm per square metre [mm2/m2]
    DL_PA_PER_KPA    : REAL := 1000.0;    // 帕到千帕的折算 [Pa/kPa] / Pascals per kilopascal [Pa/kPa]
    DL_TWO           : REAL := 2.0;       // 孔口出流式的系数 2 [-] / Orifice equation factor 2 [-]
    DL_SEC_PER_H     : REAL := 3600.0;    // 小时到秒的时基折算 [s/h] / Seconds per hour [s/h]
    DL_COEF_HI       : REAL := 1.0;       // 流量系数物理上限 [-]/ Discharge coefficient upper bound [-]
    DL_FLOW_HI_M3H   : REAL := 10000.0;   // 流量量级闸上限 [m3/h] / Flow magnitude upper bound [m3/h]
END_VAR

(* —— 段 1：非有限值闸（R19：闸断实值通路） —— *)
IF NOT (fNozzleDiaMm > -DL_BIG AND fNozzleDiaMm < DL_BIG)
   OR NOT (fPumpPressKpa > -DL_BIG AND fPumpPressKpa < DL_BIG)
   OR NOT (fDensityKgm3 > -DL_BIG AND fDensityKgm3 < DL_BIG)
   OR NOT (fDischCoef > -DL_BIG AND fDischCoef < DL_BIG)
   OR NOT (fFlowMaxM3h > -DL_BIG AND fFlowMaxM3h < DL_BIG) THEN
    fFlowM3h := 0.0;                        // 输出强制 0.0，切断污染源 / Force zero, cut polluted path
    fVelMs := 0.0;                          // 流速强制 0.0 / Velocity forced to zero
    fNozzleAreaMm2 := 0.0;                  // 面积强制 0.0 / Area forced to zero
    xFlowOver := FALSE;                     // 失效侧超限位保持假 / Overrun stays false
    xValid := FALSE;                        // 有效位清零 / Validity cleared
    FC_DL_OverflowDyeFlowCalc := FALSE;     // 返回码与有效位同源 / Return mirrors validity
    RETURN;                                 // 立即退出 / Immediate exit
END_IF

(* —— 段 2：孔径/密度零闸与系数域闸（面积为孔径平方乘子，密度为根号分母） —— *)
IF (fNozzleDiaMm <= DL_EPS)                                       // 孔径不可为零
   OR (fDensityKgm3 <= DL_EPS)                                    // 密度不可为零
   OR (fDischCoef <= 0.0)                                         // 流量系数必须为正
   OR (fDischCoef > DL_COEF_HI)                                   // 流量系数不得大于 1
   OR (nNozzle < 1)                                               // 喷嘴数至少一个
   OR (fPumpPressKpa < 0.0)                                       // 压差不得为负（根号内不可为负）
   OR (fFlowMaxM3h <= DL_EPS) THEN                                // 流量上限必须已组态
    fFlowM3h := 0.0;                        // 参数不可用即无流量 / No parameter, no flow
    fVelMs := 0.0;                          // 流速不可算 / Velocity not computable
    fNozzleAreaMm2 := 0.0;                  // 面积不可算 / Area not computable
    xFlowOver := FALSE;                     // 超限位保持假 / Overrun stays false
    xValid := FALSE;                        // 判无效 / Invalid
    FC_DL_OverflowDyeFlowCalc := FALSE;     // 返回码同步 / Return synchronised
    RETURN;                                 // 提前退出 / Early exit
END_IF

(* —— 段 3：主算式（不钳制，先出原始值供段 4 判据使用，R24） —— *)
_fAreaOneM2 := DL_PI * DL_QUARTER * fNozzleDiaMm * fNozzleDiaMm / DL_MM2_PER_M2;   // 单孔面积 [m2]
_fAreaTotalM2 := _fAreaOneM2 * INT_TO_REAL(nNozzle);                              // 总开孔面积 [m2]
_fPressPa := fPumpPressKpa * DL_PA_PER_KPA;                                       // 泵压 [Pa]
_fVelRawMs := SQRT(DL_TWO * _fPressPa / fDensityKgm3);                            // 出口流速 [m/s]
_fFlowRawM3s := fDischCoef * _fAreaTotalM2 * _fVelRawMs;                          // 流量 [m3/s]
_fFlowRawM3h := _fFlowRawM3s * DL_SEC_PER_H;                                      // 流量 [m3/h]
fNozzleAreaMm2 := _fAreaTotalM2 * DL_MM2_PER_M2;                                  // 总开孔面积 [mm2]

(* —— 段 4：判据（取原始值；单点 BOOL 聚合避免多处赋 FALSE 覆盖） —— *)
xFlowOver := (_fFlowRawM3h > fFlowMaxM3h);                                        // 流量越上限
xValid := (_fVelRawMs >= 0.0)                                                     // 流速不得为负（开方恒非负）
          AND (_fFlowRawM3h >= 0.0)                                               // 流量不得为负
          AND (_fFlowRawM3h <= DL_FLOW_HI_M3H)                                    // 不超量级闸上限
          AND (fFlowMaxM3h <= DL_FLOW_HI_M3H);                                    // 上限须在量级闸内

(* —— 段 5：输出单点写盘（钳制到物理域内，判定结果已在段 4 定案） —— *)
fFlowM3h := LIMIT(0.0, _fFlowRawM3h, fFlowMaxM3h);                                // 流量钳 0..工艺上限 [m3/h]
fVelMs := LIMIT(0.0, _fVelRawMs, DL_FLOW_HI_M3H);                                 // 流速钳物理域 [m/s]
FC_DL_OverflowDyeFlowCalc := xValid;                                              // 返回码：TRUE = 计算可信

END_FUNCTION

(* ---- FC_DL_PackedBedHtu.st ---- *)
(*
  道莅工业代码库 / Daoli Industrial ST Library
  组件: FC_DL_PackedBedHtu
  分类: DL_Process
  开源溯源: 无（clean-room 工程公式自研；参考公开工艺计算公式，未复制任何受版权保护代码）
  许可证: 本项目自有 (MIT)
  功能: 填料吸收塔传质单元高度 HTU 与塔高估算（含 1.2 倍设计余量）
  假设声明: 气相摩尔质量按空气口径 29 kg/kmol 折算 kmol/h（低浓度污染物可忽略）
*)
FUNCTION FC_DL_PackedBedHtu : BOOL
VAR_INPUT
    rGasKgH : REAL; // 气相质量流量 [kg/h] / gas mass flow
    rLiquidKgH : REAL; // 液相质量流量 [kg/h] / liquid mass flow
    rKgaKmolM3h : REAL; // 体积总传质系数 Kga [kmol/(m3·h·atm)] / overall volumetric mass transfer coefficient
    rAreaM2 : REAL; // 塔截面积 [m2] / column cross-section area
    rNtu : REAL; // 传质单元数 NTU [-] / number of transfer units
    rPressAtm : REAL; // 操作压力 [atm]，Kga 为 atm 基 / operating pressure, Kga basis
END_VAR
VAR_OUTPUT
    rHtuM : REAL; // 传质单元高度 [m] / height of a transfer unit
    rHeightM : REAL; // 填料层高度（含余量）[m] / packed bed height with margin
    bValid : BOOL; // 结果有效位 [-] / result valid flag
    iErrCode : INT; // 事件码 0=正常 1=Kga 非法 2=塔截面非法 3=无液相（填料未润湿）4=NTU 非法 5=结果非有限 / event code
END_VAR
VAR CONSTANT
    rMolWtGas : REAL := 29.0; // 气相平均摩尔质量 [kg/kmol] / mean gas molar mass
    rHeightMargin : REAL := 1.2; // 塔高设计余量系数 [-] / packed height design margin
END_VAR
VAR
    rGasKmolH : REAL; // 气相摩尔流量 [kmol/h] / gas molar flow
    rHtuRaw : REAL; // 未校验 HTU [m] / unchecked HTU
END_VAR

    // —— 段 0：全路径预清 —— //
    rGasKmolH := 0.0;
    rHtuRaw := 0.0;
    rHtuM := 0.0;
    rHeightM := 0.0;
    bValid := FALSE;
    iErrCode := 0;
    FC_DL_PackedBedHtu := FALSE;
    // —— 段 1：分母闸（传质系数、塔截面） —— //
    IF rKgaKmolM3h <= 0.0 THEN
        iErrCode := 1; // 传质系数非法，HTU 无定义 / invalid mass transfer coefficient
        RETURN;
    END_IF;
    IF rAreaM2 <= 0.0 THEN
        iErrCode := 2; // 塔截面非法 / invalid column area
        RETURN;
    END_IF;
    // —— 段 2：液相存在性闸（无液膜则 Kga 不成立） —— //
    IF rLiquidKgH <= 0.0 THEN
        iErrCode := 3; // 无液相，填料未润湿，Kga 无效 / no liquid, packing not wetted, Kga invalid
        RETURN;
    END_IF;
    IF rNtu <= 0.0 THEN
        iErrCode := 4; // NTU 非法，塔高无意义 / invalid NTU
        RETURN;
    END_IF;
    // —— 段 3：量纲链 (kg/h)/(kg/kmol) = kmol/h；/(kmol/(m3·h)·m2) = m —— //
    rGasKmolH := rGasKgH / rMolWtGas; // 气相摩尔流量 [kmol/h] / gas molar flow
    // Kga 以 atm 为基准，故分母必须乘操作压力；漏乘 P 会把 HTU 高估 P 倍
    // 量纲: (kmol/h) / (kmol/(m3·h·atm) × m2 × atm) = m
    rHtuRaw := rGasKmolH / (rKgaKmolM3h * rAreaM2 * rPressAtm); // HTU [m] / height of transfer unit
    IF ABS(rHtuRaw) > 1.0E15 THEN
        iErrCode := 5; // 结果非有限，强制归零 / non-finite result, forced to zero
        RETURN;
    END_IF;
    IF rHtuRaw < 0.0 THEN
        rHtuM := 0.0; // 负流量防御 / negative flow guard
    ELSE
        rHtuM := rHtuRaw;
    END_IF;
    // —— 段 4：塔高 = HTU × NTU × 余量（量纲 m×-×- = m） —— //
    rHeightM := rHtuM * rNtu * rHeightMargin; // 填料层高度 [m] / packed height
    bValid := TRUE;
    FC_DL_PackedBedHtu := TRUE;
END_FUNCTION
